(* Logix 5000 project; controller TFF vendor 1 type 14 code 107 rev 34.11; software revision 34.03 *)
// Mobius FlexReady

TASK HighPriority (periodic, rate 25 ms, priority 1, watchdog 2000 ms) : MainProgram   // High Priority Task
TASK MainTask (continuous, watchdog 500 ms) : Process, CCPSystem
TASK Task5ms (periodic, rate 5 ms, priority 10, watchdog 500 ms) : MainProgram5ms

MODULES
   Local : vendor 1 type 14 code 107 (Compact 0, rev 34.11)
      RACK_MURR_NODE1_TF3S : ETHERNET-MODULE (Ethernet 10.20.56.124, rev 1.1, Output RPI 5 ms)
      RACK_MURR_NODE5_TANK100 : ETHERNET-MODULE (Ethernet 10.20.56.162, rev 1.1, Output RPI 10 ms)
      RACK_MURR_NODE7_IND131_WI101 : ETHERNET-MODULE (Ethernet 10.20.56.141, rev 1.1, Output RPI 50 ms)
           RACK_MURR_NODE7_IND131_WI101:I.Data[1].15   // Data OK
           RACK_MURR_NODE7_IND131_WI101:I.Data[1]   // Slot 1 Scale Status
           RACK_MURR_NODE7_IND131_WI101:I.Data[0]   // Slot 1 Weight Data
           RACK_MURR_NODE7_IND131_WI101:O.Data[0]   // Slot 1 Tare/Target Value
           RACK_MURR_NODE7_IND131_WI101:O.Data[1]   // IND131 Command word Select weight display in net mode Clear all cmd excepted Tare and zero
      RACK_MURR_NODE0_SMART : ETHERNET-MODULE (Ethernet 10.20.56.131, rev 1.1, Output RPI 10 ms)
      RACK_MURR_NODE1_TF2S : ETHERNET-MODULE (Ethernet 10.20.56.123, rev 1.1, Output RPI 5 ms)
      RACK_MURR_NODE3_PUMP : ETHERNET-MODULE (Ethernet 10.20.56.151, rev 1.1, Output RPI 10 ms)
      RACK_MURR_NODE4_INSTRUM_TFF1 : ETHERNET-MODULE (Ethernet 10.20.56.172, rev 1.1, Output RPI 10 ms)
      RACK_MURR_NODE4_INSTRUM_TFF2 : ETHERNET-MODULE (Ethernet 10.20.56.173, rev 1.1, Output RPI 10 ms)
      RACK_MURR_NODE4_INSTRUM_TFF3 : ETHERNET-MODULE (Ethernet 10.20.56.174, rev 1.1, Output RPI 10 ms)
      RACK_MURR_NODE4_INSTRUM_TFF4 : ETHERNET-MODULE (Ethernet 10.20.56.175, rev 1.1, Output RPI 10 ms)
      RACK_MURR_NODE4_INSTRUM_TFF5 : ETHERNET-MODULE (Ethernet 10.20.56.176, rev 1.1, Output RPI 10 ms)
      RACK_MURR_NODE5_TANK250 : ETHERNET-MODULE (Ethernet 10.20.56.163, rev 1.1, Output RPI 10 ms)
      RACK_MURR_NODE5_TANK50 : ETHERNET-MODULE (Ethernet 10.20.56.161, rev 1.1, Output RPI 10 ms)
      RACK_MURR_NODE6_IND331_WI001 : ETHERNET-MODULE (Ethernet 10.20.56.142, rev 1.1, Output RPI 50 ms)
           RACK_MURR_NODE6_IND331_WI001:I.Data[1].15   // Data OK
           RACK_MURR_NODE6_IND331_WI001:I.Data[1]   // Slot 1 Scale Status
           RACK_MURR_NODE6_IND331_WI001:I.Data[0]   // Slot 1 Weight Data
           RACK_MURR_NODE6_IND331_WI001:O.Data[0]   // Slot 1 Tare/Target Value
           RACK_MURR_NODE6_IND331_WI001:O.Data[1]   // IND331 Command word Select weight display in net mode Clear all cmd excepted Tare and zero
END_MODULES

TYPE AlarmAnalog :   // Analog Alarm UDT
STRUCT
   Override : BOOL;   // Alarm Override
   Disable : BOOL;   // Alarm Disabled
   LOLOAlarm : BOOL;   // LOLO Alarm Condition
   LOAlarm : BOOL;   // LO Alarm Condition
   HIAlarm : BOOL;   // HI Alarm Condition
   HIHIAlarm : BOOL;   // HIHI Alarm Condition
   LOLODisable : BOOL;   // LOLO Alarm Disable
   LODisable : BOOL;   // LO Alarm Disable
   HIDisable : BOOL;   // HI Alarm Disable
   HIHIDisable : BOOL;   // HIHI Alarm Disable
   LOLOAck : BOOL;   // LOLO Alarm Acknowledged
   LOAck : BOOL;   // LO Alarm Acknowledged
   HIAck : BOOL;   // HI Alarm Acknowledged
   HIHIAck : BOOL;   // HIHI Alarm Acknowledged
   HIHIEnable : BOOL;   // HIHI Alarm Always Enabled for Critical Safety Alarms
   FeedPumpEnable : BOOL;   // LOLO and LO Alarm conditionned on Feed Pump Enable
   TransferPumpEnable : BOOL;   // LOLO and LO Alarm conditionned on Transfer Pump Enable
   LOLOAlarmONS : BOOL;   // Saves last value of alarm
   LOAlarmONS : BOOL;   // Saves last value of alarm
   HIAlarmONS : BOOL;   // Saves last value of alarm
   HIHIAlarmONS : BOOL;   // Saves last value of alarm
   FeedPumpTag : DINT;   // Feed Pump Tag for Pump Enable function
   TransferPumpTag : DINT;   // Transfer Pump Tag for Pump Enable function
   Value : DINT;   // Alarm Value : 0= No Alarm. 1=Non-Critical. 2= Non-Critical Unacknowledged. 3=Critical. 4=Critical Unacknowledged.
   ValueHMI : DINT;   // Alarm Value for HMI: 0= No Alarm. 1=Non-Critical. 2= Non-Critical Unacknowledged. 3=Critical. 4=Critical Unacknowledged.
   LOLO : REAL;   // LOLO Alarm Set Point
   LO : REAL;   // LO Alarm Set Point
   HI : REAL;   // HI Alarm Set Point
   HIHI : REAL;   // HIHI Alarm Set Point
   PV : REAL;   // Process Variable Value
   LOLOTimer : TIMER;   // LOLO Alarm Timer
   LOLOTimerSP : DINT;   // LOLO Alarm Timer setpoint (sec)
   LOTimer : TIMER;   // LO Alarm Timer
   LOTimerSP : DINT;   // LO Alarm Timer setpoint (sec)
   HITimer : TIMER;   // HI Alarm Timer
   HITimerSP : DINT;   // HI Alarm Timer setpoint (sec)
   HIHITimer : TIMER;   // HIHI Alarm Timer
   HIHITimerSP : DINT;   // HIHI Alarm Timer setpoint (sec)
   EnableCfg : BOOL;   // Set to 1 to Configure \ Use Analog Alarm
END_STRUCT
END_TYPE

TYPE AlarmControl :   // Alarm Control UDT
STRUCT
   DESC : STRING25;   // Description
   EGU : STRING5;   // Unit
   AlarmAck : BOOL;   // Alarm Acknowledge Flag
   AlarmHigh : BOOL;   // Critical Alarm Condition
   AlarmLow : BOOL;   // Non-Critical Alarm Condition
   AlarmHighUnack : BOOL;   // Critical Unacknowledged Alarm Condition
   AlarmLowUnack : BOOL;   // Non-Critical Unacknowledged Alarm Condition
   HighHMI : BOOL;   // Critical Alarm Condition (for HMI)
   LowHMI : BOOL;   // Non-Critical Alarm Condition (for HMI)
   HighUnackHMI : BOOL;   // Critical Unacknowledged Alarm Condition (for HMI)
   LowUnackHMI : BOOL;   // Non-Critical Unacknowledged Alarm Condition (for HMI)
   Horn : BOOL;   // Alarm Horn
   YellowLamp : BOOL;   // Non-Critical Alarm Indicator
   RedLamp : BOOL;   // Critical Alarm Indicator
   Current : BOOL;   // Current Alarm Status
   AckOutput : BOOL;   // Alarm Acknowledge Output
   FlashControl : BOOL;   // Flash Control
   EnableAllIn : BOOL;   // Enable All Alarms Input
   EnableAllOut : BOOL;   // Enable All Alarms Output
   DisableAllIn : BOOL;   // Disable All Alarms Input
   DisableAllOut : BOOL;   // Disable All Alarms Output
   NewAlarm : BOOL;   // True for 1 scan when new alarm is detected
   SilenceHorn : BOOL;   // Set true to Silence horn
   FlashTimer : TIMER;   // Flash Timer
   AckTimer : TIMER;   // Acknowledge Timer
   EnableAllTimer : TIMER;   // Enable All Alarms Timer
   DisableAllTimer : TIMER;   // Disable All Alarms Timer
   HornAddress : INT;   // Output address for Alarm horn
   EnableAllAnaSigIn : BOOL;   // Enable All analog signal failure Alarms Input
   EnableAllAnaSigOut : BOOL;   // Enable All analog signal failure Alarms Output
   DisableAllAnaSigIn : BOOL;   // Disable All analog signal failure Alarms Input
   DisableAllAnaSigOut : BOOL;   // Disable All analog signal failure Alarms Output
   EnableAllAnaSigTimer : TIMER;   // Enable All analog signal failure Alarms Timer
   DisableAllAnaSigTimer : TIMER;   // Disable All analog signal failure Alarms Timer
   AlarmHighMem : BOOL;   // Critical Alarm Condition Mem
   ESAckAddress : INT;   // Output address for re-established system
   ESAckTimer : TIMER;   // Emergency Stop Acknowledge Timer
   ESAck : BOOL;   // Emergency Stop Acknowledge
   InitAlarmConfig : BOOL;   // Initialize alarms config if the command is set from the HMI
END_STRUCT
END_TYPE

TYPE AlarmDeviation :   // Deviation Alarm UDT
STRUCT
   Override : BOOL;   // Alarm Override
   Disable : BOOL;   // Alarm Disabled
   HIAlarm : BOOL;   // HI Deviation Alarm Condition
   HIHIAlarm : BOOL;   // HIHI Deviation Alarm Condition
   HIDisable : BOOL;   // HI Alarm Disable
   HIHIDisable : BOOL;   // HIHI Alarm Disable
   HIAck : BOOL;   // HI Alarm Acknowledged
   HIHIAck : BOOL;   // HIHI Alarm Acknowledged
   LOLOAlarmONS : BOOL;   // One shot when alarm occures
   HIAlarmONS : BOOL;   // One shot when alarm occures
   LOAlarmONS : BOOL;   // One shot when alarm occures
   HIHIAlarmONS : BOOL;   // One shot when alarm occures
   Value : DINT;   // Alarm Value
   ValueHMI : DINT;   // Alarm Value for HMI
   HI : REAL;   // HI Alarm Set Point
   HIHI : REAL;   // HIHI Alarm Set Point
   LOLOLim : REAL;   // LOLO Alarm Set Point (calculated)
   LOLim : REAL;   // LO Alarm Set Point (calculated)
   HILim : REAL;   // HI Alarm Set Point (calculated)
   HIHILim : REAL;   // HIHI Alarm Set Point (calculated)
   HITimer : TIMER;   // HI Alarm Timer
   HITimerSP : DINT;   // HI Alarm Timer setpoint (sec)
   HIHITimer : TIMER;   // HIHI Alarm Timer
   HIHITImerSP : DINT;   // HIHI Alarm Timer setpoint (sec)
   EnableCfg : BOOL;   // Set to enable alarm
END_STRUCT
END_TYPE

TYPE AnalogInput :   // Analog Input UDT
STRUCT
   TagName : STRING6;   // PID Tag Name
   TagDisplayName : STRING6;   // PID Tag Name
   OutofRange : BOOL;   // Out of Range
   FilterType : BOOL;   // Filter Type 0=LP, 1=Avg
   AveragingTotal : DINT;   // Averaging Filter Total
   Address : DINT;   // Input Address (RawAnalogInputArray)
   RawMin : DINT;   // Raw Minimum Range
   RawMax : DINT;   // Raw Maximum Range
   RawValue : DINT;   // Raw Value (Measuring value given by the I/O card)
   RawLowLimit : DINT;   // Raw Out of Range LO Limit
   RawHighLimit : DINT;   // Raw Out of Range HI Limit
   FilterUser : DINT;   // User Filter Value
   FilteredRaw : DINT;   // Raw Filtered Value
   FilterActual : REAL;   // Actual Filter Value
   ScaledMin : REAL;   // Scaled Minimum Range
   ScaledMax : REAL;   // Scaled Maximum Range
   CurrentValue : REAL;   // Current Value
   RangeMin : REAL;   // Scaled Minimum Range (Config Analog Points)
   RangeMax : REAL;   // Scaled Maximum Range (Config Analog Points)
   RangeMinSave : REAL;   // Scaled Minimum Range (previous)
   RangeMaxSave : REAL;   // Scaled Maximum Range (previous)
   RealCfg : BOOL;   // Set to 1 if real analog input is used. Set to 0 for soft input (derived data)
   EnableCfg : BOOL;   // Set to 1 to activate this Tag
   OverrideCfg : BOOL;   // Set to 1 to allow user to Overide alarm
   Desc : STRING25;   // Description
   EGU : STRING5;   // Unit
END_STRUCT
END_TYPE

TYPE AnalogOutput :   // Analog Output UDT
STRUCT
   Tag : STRING10;   // Tag name
   RawValue : DINT;   // Raw Value Send to I/O Card
   RawMin : DINT;   // Raw Min
   RawMax : DINT;   // Raw Max
   ScaledValue : REAL;   // Scaled Value
   ScaledMin : REAL;   // Scaled Minimum Range
   ScaledMax : REAL;   // Scaled Maximum Range
   EnableCfg : BOOL;   // Set to 1 to enable Analog Output
END_STRUCT
END_TYPE

TYPE AverageCalculation :
STRUCT
   SUM : REAL;   // Sum of average
   COUNTER : DINT;   // Counter of average
   TIMER : TIMER;   // Timer of average
   TIMER_OSR : BOOL;   // Timer one shot
END_STRUCT
END_TYPE

TYPE CCPSystem :   // CCP System UDT
STRUCT
   Run : BOOL;   // Run Flag
   RunAuto : BOOL;   // Auto Run Flag
   Procedure : BOOL;   // Procedure Flag
   Complete : BOOL;   // Procedure Complete
   Download : BOOL;   // Manual Download
   Heartbeat : BOOL;   // CCPRuntime Heartbeat
   OperationDownloadFlag : BOOL;   // Legacy Tag. Not used by PLC
   OperationStartFlag : BOOL;   // Operation Start Flag
   Manual : BOOL;   // Recipe Pool Flag
   State : DINT;   // Machine State
   Language : DINT;   // Language Number
   ErrorPhase : DINT;   // Error in Phase #
   ErrorStep : DINT;   // Error in Step #
   Error : DINT;   // Error Description
   OperationNoInBatch : DINT;   // Legacy Tag. Not used by PLC
   EndPointer : DINT;   // End Operation Step Buffer Pointer
   Machine : STRING;   // Machine Name
   ProductID : STRING;   // Batch Product ID from Operation Header
   Description : STRING;   // Batch Description from Operation Header
   Created : STRING;   // Date and Time when the last operation has been downloaded in PLC
   Originator : STRING;   // Last saved by field from Operation Header
   Comment : STRING;   // Comment
   OperationName : STRING90;   // Name and path of last operation downloaded in PLC
   ConfigFile : STRING;   // Current configuration file used
   LastMod : STRING;   // Last Mod
   GradientBasis : STRING;   // Gradient Basis
   GradientVariable : STRING;   // Gradient Variable
   GradientSegments : STRING;   // Gradient Segments
   StateWatchDog : TIMER;   // If Downloading for longer than this time the state will reset to 0
   EventList : EventList;   // Event List Array
   BufferSteps : STRING25[251];   // Buffer Steps Array
   BufferEvents : STRING50[251];   // Buffer Events Array
   HETP_ON_OFF : BOOL;   // HETP (1 = Start , 0 = Stop)
   DefaultOnComplete : BOOL;   // At the end of recipe apply default flowpath (0 = Apply , 1 = Don't Apply)
END_STRUCT
END_TYPE

TYPE CCPSystem_Storage :
STRUCT
   Run : BOOL;   // Run Flag
   RunAuto : BOOL;   // Auto Run Flag
   Procedure : BOOL;   // Procedure Flag
   Complete : BOOL;   // Procedure Complete
   Download : BOOL;   // Manual Download
   Heartbeat : BOOL;   // CCPRuntime Heartbeat
   OperationDownloadFlag : BOOL;   // Legacy Tag. Not used by PLC
   OperationStartFlag : BOOL;   // Operation Start Flag
   TestAction : BOOL;   // Action Test Flag
   Manual : BOOL;   // Recipe Pool Flag
   State : DINT;   // Machine State
   Language : DINT;   // Language Number
   ErrorPhase : DINT;   // Error in Phase #
   ErrorStep : DINT;   // Error in Step #
   Error : DINT;   // Error Description
   OperationNoInBatch : DINT;   // Legacy Tag. Not used by PLC
   EndPointer : DINT;   // End Operation Step Buffer Pointer
   Machine : STRING;
   ProductID : STRING;
   Description : STRING;
   Created : STRING;
   Originator : STRING;
   Comment : STRING;
   OperationName : STRING90;
   ConfigFile : STRING;
   LastMod : STRING;
   GradientBasis : STRING;
   GradientVariable : STRING;
   GradientSegments : STRING;
   StateWatchDog : TIMER;   // If Downloading for longer than this time the state will reset to 0
END_STRUCT
END_TYPE

TYPE ChartMark :   // Chart Mark UDT
STRUCT
   In : BOOL;   // Chart Mark In
   Out : BOOL;   // Chart Mark Out
END_STRUCT
END_TYPE

TYPE Concentration :   // Concentration UDT
STRUCT
   VCF : REAL;   // Volume Concentration Factor
   CB : REAL;   // Protein Concentration
   Conc_Init : REAL;   // Initial Protein Concentration SP
   Conc_Final : REAL;   // Final Protein Concentration SP
   Conc_Final_Volume : REAL;   // Final Concentration Volume SP
   Final_Conc_Volume_Reached : BOOL;   // Final Concentration Volume Reached
   Final_Conc_Volume_DownTimer : TIMER;   // Final Concentration Volume Deactivation timer
   Final_Conc_Volume_UpTimer : TIMER;   // Final Concentration Volume Activation timer
   Final_Conc_Protein_Reached : BOOL;   // Final Protein Concentration Reached
   Final_Conc_Protein_DownTimer : TIMER;   // Final Protein Concentration Deactivation timer
   Final_Conc_Protein_UpTimer : TIMER;   // Final Protein Concentration Activation timer
   LogConcIn : BOOL;   // Log Concentration Input
   LogConcOut : BOOL;   // Log Concentration Output
   LogConcTimer : TIMER;   // Log Concentation Timer
END_STRUCT
END_TYPE

TYPE Configuration :   // Configuration UDT
STRUCT
   Reset : BOOL;   // Activate Reset Loop Configuration
   IndexA0 : DINT;   // Index AnalogOutput
   IndexAP : DINT;   // Index AnalogPoint
   IndexDP : DINT;   // Index DigitalPoint
   IndexDr : DINT;   // Index Drive
   IndeXValve : DINT;   // Index Valve
   IndexReset : DINT;   // Index Reset
   IndexCL : DINT;   // Index Control Loop
   IndexFlowpath : DINT;   // Index Flowpath
END_STRUCT
END_TYPE

TYPE ControlLoop :   // Control Loop UDT
STRUCT
   Tag : STRING5;   // Tag Name
   Desc : STRING25;   // Description
   LoopCfg : BOOL;   // Set to 1 to use this loop
   ManualEGU : STRING5;   // Unit of Manual Control Mode
   AutoEGU : STRING5;   // Unit of Auto Control Mode
   Auto1EGU : STRING5;   // Unit of Auto Control Mode 1
   Auto2EGU : STRING5;   // Unit of Auto Control Mode 2
   Auto3EGU : STRING5;   // Unit of Auto Control Mode 3
   Interlock : BOOL;   // Loop Interlock
   Enable : BOOL;   // Loop Enabled
   Manual : BOOL;   // Control Mode 0=Auto, 1=Manual
   Stable : BOOL;   // Loop Stable
   DBOK : BOOL;   // Control Within Deadband
   Status : INT;   // Status
   Auto1 : BOOL;   // Auto Control Mode 1
   Auto2 : BOOL;   // Auto Control Mode 2
   Auto3 : BOOL;   // Auto Control Mode 3
   Auto4 : BOOL;   // Auto Control Mode 4
   StepUp : BOOL;   // Increment CV
   StepDown : BOOL;   // Decrement CV
   RampEnable : BOOL;   // Ramp Enable
   RampUp : BOOL;   // Ramping UP
   RampDown : BOOL;   // Ramping Down
   RampStatus : BOOL;   // Ramping Status
   RampAutoOSR : BOOL;   // Auto Ramp One-Shot
   RampManualOSR : BOOL;   // Manual Ramp One-Shot
   PIDEnable : BOOL;   // PID Enabled
   ManualOSR : BOOL;   // Manual Mode One-Shot
   Auto1OSR : BOOL;   // Control Mode 1 One-Shot
   Auto2OSR : BOOL;   // Control Mode 2 One-Shot
   Auto3OSR : BOOL;   // Control Mode 3 One-Shot
   Auto4OSR : BOOL;   // Control Mode 4 One-Shot
   StepIncrement : DINT;   // Step Increment/Decrement Value
   CycleTime : DINT;   // Cycle Time (for modulating output)
   PV : REAL;   // Process Variable
   PVAuto1 : REAL;   // Process Variable for Control Mode Auto 1
   PVAuto2 : REAL;   // Process Variable for Control Mode Auto 2
   PVAuto3 : REAL;   // Process Variable for Control Mode Auto 3
   PVAuto4 : REAL;   // Process Variable for Control Mode Auto 4
   CV : REAL;   // Control Value
   SPAuto : REAL;   // Auto Set Point
   SPAutoSave : REAL;   // Auto Set Point (previous)
   SPAuto1 : REAL;   // Auto Set Point Mode 1
   SPAuto2 : REAL;   // Auto Set Point Mode 2
   SPAuto3 : REAL;   // Auto Set Point Mode 3
   SPAuto4 : REAL;   // Auto Set Point Mode 4
   SPManual : REAL;   // Manual Set Point
   SPManualSave : REAL;   // Manual Set Point (previous)
   RangeMin : REAL;   // Min EGU Range
   RangeMax : REAL;   // Max EGU Range
   SPRangeMin : REAL;   // Set Point Min EGU Range
   SPRangeMax : REAL;   // Set Point Max EGU Range
   RampRate : REAL;   // Ramp Rate
   RampRateSave : REAL;   // Ramp Rate (previous)
   RampStart : REAL;   // Ramp Start Value
   Deadband : REAL;   // Deadband
   DBLO : REAL;   // Low Deadband Value
   DBHI : REAL;   // High Deadband Value
   RampTimer : TIMER;   // Ramp Timer
   StableTimer : TIMER;   // Loop Stable Timer
   StableTime : DINT;   // Loop Stable Time setpoint (sec)
   PIDTimer : TIMER;   // PID Timer
   CycleTimer : TIMER;   // Cycle Timer (for modulating output)
   PID : PID;   // PID Instruction Data
   KP : REAL[3];   // Loop Gain from HMI
   KI : REAL[3];   // Loop Reset from HMI
   KD : REAL[3];   // Loop Rate from HMI
   DB : REAL[3];   // Loop Deadband from HMI
   On : BOOL;   // Turns all controll On
   DisOSR : BOOL;   // One Shot DisOSR
   OutputOn_OSR : BOOL;   // One Shot OutputOn_OSR
   OutputOff_OSR : BOOL;   // One Shot OutputOff_OSR
   DigitalOutput : BOOL;   // Output from loop in for descrete control
   RampCfg : BOOL;   // Set to 1 to Enable Ramp Option
   Auto1Cfg : BOOL;   // Set to 1 to use Auto 1 option
   Auto2Cfg : BOOL;   // Set to 1 to use Auto 2 option
   Auto3Cfg : BOOL;   // Set to 1 to use Auto 3 option
   Auto4Cfg : BOOL;   // Set to 1 to use Auto 4 option
   Auto1PVCfg : DINT;   // Set to Analog Point Number
   Auto2PVCfg : DINT;   // Set to Analog Point Number
   Auto3PVCfg : DINT;   // Set to Analog Point Number
   Auto4PVCfg : DINT;   // Set to Analog Point Number
   Auto1RangeMax : REAL;   // Set Point EGU Range Max
   Auto2RangeMax : REAL;   // Set Point EGU Range Max
   Auto3RangeMax : REAL;   // Set Point EGU Range Max
   Auto4RangeMax : REAL;   // Set Point EGU Range Max
   AutoSwitchEnable : BOOL;   // Set to 1 to allow loop to switch from auto1 to auto 2
   OutputAddress : INT;   // Set to analog output to use for this loop
   LoopStatus : INT;   // Loop Mode Status for HMI
END_STRUCT
END_TYPE

TYPE CriteriaFlag :   // Criteria Flag UDT
STRUCT
   Flag1 : BOOL;   // Criteria Flag 1 (1=ON , 0=OFF)
   Flag2 : BOOL;   // Criteria Flag 2 (1=ON , 0=OFF)
   Flag3 : BOOL;   // Criteria Flag 3 (1=ON , 0=OFF)
   Flag4 : BOOL;   // Criteria Flag 4 (1=ON , 0=OFF)
   Flag5 : BOOL;   // Criteria Flag 5 (1=ON , 0=OFF)
END_STRUCT
END_TYPE

TYPE CVTune :   // Control Valve Tuning Data Type
STRUCT
   ClosedRaw : REAL;   // Captured Raw Value When Valve is Closed
   OpenRaw : REAL;   // Captured Raw Value When Valve is Open
   MinOutput : REAL;   // Minimum output for tuning adjustment for valve
   MaxOutput : REAL;   // Maximum output for tuning adjustment for valve
   MinTimer : TIMER;   // Timer to capture closed raw value
   MaxTimer : TIMER;   // Timer to capture open raw value
   OSR : INT;   // One shot bits
   Activate : BOOL;   // Activate tuning function
   Enable : BOOL;   // Tuning routine is enabled
END_STRUCT
END_TYPE

TYPE DCS :
STRUCT
   ActionsParameters : DCSParameters;   // Recipe Parameters
   Criteria : DCSCriteria;   // Recipe Criteria
   RunCmd : BOOL;   // Start Recipe Command
   ShowHeader : BOOL;   // Show Pre and Post Run Header
   RunID : STRING50;   // Recipe Header Run ID (Must be unique)
   UserName : STRING80;   // Recipe Header User Name
   ProductID : STRING80;   // Recipe Header Product ID
   BatchID : STRING80;   // Recipe Header Batch ID
   StepID : STRING80;   // Recipe Header Step ID
   FileName : STRING240;   // File Name for Start recipe (if not using RecipePoolID)
   PreRunComment : STRING240;   // Recipe Header Pre Run Comment
   PostRunComment : STRING240;   // Recipe Header Post Run Comment
   RecipePoolID : DINT;   // Recipe Pool ID for Start recipe (If 0 the file name will be used)
   Status : DINT;   // System status for DCS
   ColumnInfo : STRING240;   // Recipe Header Column Info
   PackedBedInfo : STRING240;   // Recipe Header Packed Bed Info
   SampleInfo : STRING240;   // Recipe Header Sample Info
   BufferInfo : STRING240;   // Recipe Header Buffer Info
END_STRUCT
END_TYPE

TYPE DCSCriteria :
STRUCT
   Criteria_1 : BOOL;
   Criteria_2 : BOOL;
END_STRUCT
END_TYPE

TYPE DCSParameters :
STRUCT
   Feed_Pump_Speed_Setpoint : REAL[3];
   Feed_Pump_Flow_Setpoint : REAL[3];
   Feed_Pump_DP_Setpoint : REAL[3];
   Level_Pump_Speed_Setpoint : REAL[3];
   Level_Pump_Level_Setpoint : REAL[3];
   PCV001_Retentate_Position_Setpoint : REAL[3];
   PCV001_Retentate_Pressure_Setpoint : REAL[3];
   PCV001_Retentate_TMP_Setpoint : REAL[3];
   PCV101_Filtrate_Position_Setpoint : REAL[3];
   PCV101_Filtrate_Flow_Setpoint : REAL[3];
   PCV101_Filtrate_TMP_Setpoint : REAL[3];
   Mixer_Speed_Setpoint : REAL[3];
   Mixer_Auto_Min_Setpoint : REAL[3];
   Mixer_Auto_Max_Setpoint : REAL[3];
   Init_Protein_Conc : REAL[1];
   Final_Protein_Conc : REAL[1];
   Final_Protein_Volume : REAL[1];
   Holdup_Volume : REAL[1];
   Init_Diaf_Volume : REAL[1];
   Final_Diaf_Volume : REAL[1];
   Membrane_Area : REAL[1];
   Membrane_Density : REAL[1];
END_STRUCT
END_TYPE

TYPE DerivedData :   // DerivedData UDT
STRUCT
   HOLDUP : REAL;   // Holdup Volume
   PI001_PSI : REAL;   // PI001 Pressure in PSI
   PI401_PSI : REAL;   // PI401 Pressure in PSI
END_STRUCT
END_TYPE

TYPE Diafiltration :   // Diafiltration UDT
STRUCT
   Diaf_Volume : REAL;   // Diafiltration Volume
   Diaf_Init : REAL;   // Initial Diafiltration Volume SP
   Diaf_Final_Volume : REAL;   // Final Diafiltration Volume SP
   Snap : BOOL;   // Level Snapshot
   Final_Diaf_Volum_Reached : BOOL;   // Final Diafiltration Volume Reached
   Final_Diaf_Volum_DownTimer : TIMER;   // Final Diafiltration Volume Deactivation timer
   Final_Diaf_Volum_UpTimer : TIMER;   // Final Diafiltration Volume Activation timer
   Diaf_Snap_Value : REAL;   // Volume value snapped
   LogDiafIn : BOOL;   // Log Diafiltration Input
   LogDiafOut : BOOL;   // Log Diafiltration Output
   LogDiafTimer : TIMER;   // Log Diafiltration Timer
END_STRUCT
END_TYPE

TYPE DigitalPoint :   // Digital Point UDT
STRUCT
   Tag : STRING10;   // PID Tag to be Used for Display
   Desc : STRING25;   // Description to be Used for Display
   CurrentValue : BOOL;   // Current value of Tag
   AlarmCurrentValue : BOOL;   // Displays state of processed alarm input.
   AlarmAck : BOOL;   // Alarm Acknowledged
   Alarm : BOOL;   // Alarm
   Override : BOOL;   // Alarm Override
   Mimic : INT;   // Set color on HMI digital point mimic
   SoftInput : BOOL;   // Used as current value when RealInputCfg is set to 0
   Condition1 : BOOL;   // Enable Condition 1 Must be True to Enable alarm condition
   Condition2 : BOOL;   // Enable Condition 2 Must be True to Enable alarm condition
   Cond1Text : STRING;   // Condtion 1 Text
   Cond2Text : STRING;   // Condition 2 text
   DelayTimer : TIMER;   // Alarm Timer
   DelayTimerSP : DINT;   // Alarm Timer setpoint (sec)
   Priority : BOOL;   // Alarm Priority 0=Low, 1=High
   EnableCfg : BOOL;   // Set to True to configure point on system
   ActiveStateCFg : BOOL;   // Set to 0 to invert incomming state
   RealInputCfg : BOOL;   // Set to 1 to Use Hardwired Input. Set to 0 to disable Hardwired and use software condition
   InputAddressCfg : DINT;   // Set to address of hardwared input to be used on alarm
   AlarmCfg : BOOL;   // Set to 1 to Use alarm on this point
   AlarmStateCfg : BOOL;   // Set to 1 to alarm on a 0 to 1 transition. Set to zero to alarm on a 1 to 0 transition
   OverrideCfg : BOOL;   // set to 1 to allow user to Override alarm
   PriorityCfg : BOOL;   // Set to 1 to allow user to set Priority and Enable
   Cond1Cfg : BOOL;   // Set to 1 to Enable Condition
   Cond2Cfg : BOOL;   // Set to 1 to Enable Condition
   FlashingInputCfg : BOOL;   // Set to 1 for Heartbeat Style Inputs
   AlarmONS : BOOL;   // One shot when alarm occurs
END_STRUCT
END_TYPE

TYPE Drive :   // Pump Control UDT
STRUCT
   TagName : STRING10;   // Drive tag name
   Desc : STRING25;   // Drive Description
   Mode : BOOL;   // Control Mode
   ManualCommand : BOOL;   // Manual Command
   AutoCommand : BOOL;   // Auto Command
   RunCommand : BOOL;   // Run Command
   RunStatus : BOOL;   // Running Status
   RunInterlock : BOOL;   // Run Interlock
   RunInput : BOOL;   // Run Digital Input 0=No, 1=Yes
   OutputAddress : DINT;   // Run Command Output Address
   InputAddress : DINT;   // Running Input Address
   InterlockTimer : TIMER;   // Interlock Delay Timer
   RunOns : BOOL;   // Run one shot
   StopOns : BOOL;   // Stop One shot
   RunRequest : BOOL;   // Run request for auto or man mode
   Interlocked : BOOL;   // Drive is commanded to run but currently stopped by interlock
   EnableCfg : BOOL;   // Set to enable Drive
   ReverseCfg : BOOL;   // Set to enable reverse control
   Direction : BOOL;   // 0 = forward. 1 = reverse
   DirectionAddress : DINT;   // Direction Output Address
   DriveStatus : INT;   // Drive Status
   DriveLoopStatus : INT;   // Drive Loop Status
   DriveAlarmStatus : INT;   // Drive Alarm Status
   ValidFlowpath : BOOL;   // Valid flowpath flag
END_STRUCT
END_TYPE

TYPE EventList :
STRUCT
   Event : DINT[1000];   // Event List Array
   Value : REAL[1000];   // Value Array
   PreRunValue : REAL[1000];   // Pre Run Value
END_STRUCT
END_TYPE

TYPE FactorySettings :   // Factory Settings
STRUCT
   ProductName : STRING90;   // Product Name
   SerialNumber : STRING90;   // Serial Number
   ComputerName : STRING90;   // Computer Name
   ComputerDesc : STRING90;   // Computer Description
   DateFormat : STRING90;   // Date Format
   FlagUK : BOOL;   // Use UK Flag instead of US
   PCV001ClosedSP : REAL;   // PCV001 Closed Set Point
   PCV101ClosedSP : REAL;   // PCV101 Closed Set Point
END_STRUCT
END_TYPE

TYPE FaultRecordType :   // Fault Record Type UDT
STRUCT
   TimeLow : DINT;   // Lower 32 bits of the fault timestamp value
   TimeHigh : DINT;   // Upperer 32 bits of the fault timestamp value
   RecType : INT;   // Fault Type
   Code : INT;   // Unique code for the fault
   Info : DINT[8];   // Fault specific information
END_STRUCT
END_TYPE

TYPE FlowPath :   // Flow Path UDT
STRUCT
   Command : BOOL;   // Flow Path Command
   Status : BOOL;   // Flow Path Status
   FlushTruth : BOOL;   // Flush Mode Enable Truth
   DrainTruth : BOOL;   // Drain Mode Enable Truth
   FlushMask : BOOL;   // Flush Mode Enable Mask
   DrainMask : BOOL;   // Drain Mode Enable Mask
   Truth1 : DINT;   // Truth Table 1 (Valves 1-32)
   Truth2 : DINT;   // Truth Table 2 (Valves 33-64)
   Truth3 : DINT;   // Truth Table 3 (Valves 65-96)
   Truth4 : DINT;   // Truth Table 4 (Valves 97-128)
   Mask1 : DINT;   // Mask 1 (Valves 1-32)
   Mask2 : DINT;   // Mask 2 (Valves 33-64)
   Mask3 : DINT;   // Mask 3 (Valves 65-96)
   Mask4 : DINT;   // Mask 4 (Valves 97-128)
   Desc : STRING;   // Flow Path Description
END_STRUCT
END_TYPE

TYPE FlowPathControl :   // Flow Path Control UDT
STRUCT
   Flag : BOOL;   // Flow Path Command Flag
   Valve1 : DINT;   // Valve Control 1 (Valves 1-32)
   Valve2 : DINT;   // Valve Control 2 (Valves 33-64)
   Valve3 : DINT;   // Valve Control 3 (Valves 65-96)
   Valve4 : DINT;   // Valve Control 4 (Valves 97-128)
   MaxFlowPath : DINT;   // Maximum Number of Flow Paths
   Status : DINT;   // Flow Path Status
   StatusHMI : DINT;   // Flow Path Status for HMI
   Save : BOOL;   // Set to 1 to save Flowpath
   SaveStored : BOOL;   // Stored Save cmd
   Restore : BOOL;   // Set to 1 to restore flowpath
   SaveOns : BOOL;   // one shot after save
   HoldOns : BOOL;   // one shot after Hold
   FlowpathEnable : BOOL[64];   // Enable Flowpath
   FlushMode_Enabled : BOOL;   // Flush Mode Enabled
   DrainMode_Enabled : BOOL;   // Drain Mode Enabled
END_STRUCT
END_TYPE

TYPE FlowPathSetup :   // Flowpath Setup UDT
STRUCT
   Apply : BOOL;   // Apply Flow Path
   Number : DINT;   // Flow Path Number
   Prev : DINT;   // Previous Flow Path Number
   Mask_View : BOOL;   // View the Mask of selected Flowpath
   Mask_Save : BOOL;   // Save the Mask of selected Flowpath
   Truth_View : BOOL;   // View the Truth of selected Flowpath
   Truth_Save : BOOL;   // Save the Truth of selected Flowpath
   OpenAllValve : BOOL;   // Set the Flowpath 61 to Open All Valves
   CloseAllValve : BOOL;   // Set the Flowpath 62 to Close All Valves
END_STRUCT
END_TYPE

TYPE IO_Station :   // Station State UDT
STRUCT
   Node_Comm_Status_value : INT;   // Node Communication Status Value (get from status of hardware card)
   Node_Comm_Status : BOOL;   // Node Communication Status (0=Defect , 1=OK)
   Node_Internal_Defect_Status_value : INT;   // Node Internal Defect Status Value (at least one defect on the node : branch, slot, channel)
   Node_Internal_Defect_Status : BOOL;   // Node Internal Defect Status (0=Defect , 1=OK)
   Inhibition : DINT;   // Inhibit \ Uninhibit Station Module
END_STRUCT
END_TYPE

TYPE LinearGradient :   // Linear Gradient UDT
STRUCT
   Enable : BOOL;   // Linear Gradient Enable
   Hold : BOOL;   // Gradient Hold
   Segments : DINT;   // Number of Segments
   Variable : DINT;   // Gradient Variable (1=Time, 2=CVs, 3=Volume)
   Basis : DINT;   // Basis (1=Percent, 2=Conductivity)
   Segment : DINT;   // Current Segment
   State : DINT;   // Sets state of control : 0 = Disabled 1 = Running 2 = Paused
   Input : REAL;   // Input Value
   Result : REAL;   // Result
   X2 : REAL;   // Current Segment Duration
   Y1 : REAL;   // Current Start Value
   Y2 : REAL;   // Current End Value
   X : REAL[21];   // Gradient X Values (Durations)
   Y : REAL[21];   // Gradient Y Values (Set Points)
END_STRUCT
END_TYPE

TYPE LoggedValue :   // Logged Value UDT
STRUCT
   Value : REAL[8];   // Value to be logged in Audit Trail (used in Event section of configuration file)
END_STRUCT
END_TYPE

TYPE Membrane_Data :   // Membrane Data UDT
STRUCT
   Flux : REAL;   // Membrane Flux
   Area : REAL;   // Membrane Area SP
   Density : REAL;   // Density
   NWP_TCF : REAL;   // NWP Temperature correction factor
   NWP_TCF_Temp : INT;   // Temp. Temperature used in NWP calculation (INT)
   NWP_TCF_Lookup_25 : REAL[53];   // Lookup table for TCF
   AlarmStatus : INT;   // Alarm Status ( 0 = No Alarm , 1 = Non Critical Alarm , 2 = Critical Alarm )
END_STRUCT
END_TYPE

TYPE Memory_Data :   // This UDT is for putting the memory information returned by the Controller
STRUCT
   Reading_Request : BOOL;   // Request of Memory data reading
   Free_Mem_IO : DINT;   // Controler data: Free I/O Memory
   Free_Mem_DT : DINT;   // Controler data: Free Data & Logic Memory
   Free_Mem_Gen : DINT;   // Controler 1756-L55M16 only: Free Expansion Memory
   Free_Memory : DINT;   // Controler data: Total Free Memory (addition)
   Total_Mem_IO : DINT;   // Controler data: Total I/O Memory
   Total_Mem_DT : DINT;   // Controler data: Total Data & Logic Memory
   Total_Mem_Gen : DINT;   // Controler 1756-L55M16 only: Total Expansion Memory
   Total_Memory : DINT;   // Controler data: Total Memory (addition)
   Biggest_Gen_Mem_Size_Ava : DINT;   // Controler 1756-L55M16 only: Additionnal Expansion Memory
   Biggest_IO_Mem_Size_Ava : DINT;   // Controler 1756-L55M16 only: Largest contiguous block of Additionnal free Expansion Memory
   Biggest_DT_Mem_Size_Ava : DINT;   // Controler dsata: Largest contiguous block of Additionnal free Expansion Memory
   Total_Mem_DT_Real : REAL;   // Controler data: Total Data & Logic Memory
   Free_Mem_DT_Real : REAL;   // Controler data: Free Data & Logic Memory
   Used_Mem_DT_Real : REAL;   // Controler data: Used Data & Logic Memory
   Percentage_Used_DT : REAL;   // Controler data: Percentage of used Data & Logic Memory
END_STRUCT
END_TYPE

TYPE Mixer :
STRUCT
   Enable : BOOL;   // Enable Mixer Control Loop
   Mode : BOOL;   // Control Mode 0=Weight, 1=Speed
   ModeONS : BOOL;   // Manual Mode One-Shot
   SPManual : REAL;   // Manual Speed Set Point
   SPAutoMin : REAL;   // Auto Max Speed Set Point
   SPAutoMax : REAL;   // Auto Min Speed Set Point
   LevelMin : REAL;   // Minimum Level
   LevelMax : REAL;   // Maximum Level
   CV : REAL;   // Control Value
   Alarm_Reset_Cmd : BOOL;   // Alarm Reset Command
   Alarm_Reset_Cmd_Timer : TIMER;   // Alarm Reset Command Timer
END_STRUCT
END_TYPE

TYPE OperatingTime :   // Operating Time Exceeded Control
STRUCT
   DayMax : REAL;   // Setpoint for Alarm Operating Time Exceeded
   HMICtrl : BOOL;   // Control Tag Reset on launch Workspace
   TimerCtrl : TIMER;   // Timer for set tag HMICtrl
   CountPre : DINT;   // Setpoint for Alarm in sec
   Counter : DINT;   // Second Counter for Alarm
END_STRUCT
END_TYPE

TYPE Operation :   // Operation UDT
STRUCT
   Step : DINT;   // Step Number
   Criteria1 : DINT;   // Criteria 1 Code
   Criteria1Operator : DINT;   // Criteria 1 Operator
   Boolean : DINT;   // Boolean
   Criteria2 : DINT;   // Criteria 2 Code
   Criteria2Operator : DINT;   // Criteria 2 Operator
   Action : DINT;   // Action Code
   Label : DINT;   // Label
   Criteria1Value : REAL;   // Criteria 1 Value
   Criteria2Value : REAL;   // Criteria 2 Value
   ActionValue : REAL;   // Action Value
END_STRUCT
END_TYPE

TYPE Options :   // Options UDT
STRUCT
   No_Filtrate_Measurement : BOOL;   // No Filtrate Measurement
   WI101 : BOOL;   // WI101 Filtrate Weight
   WI102 : BOOL;   // WI102 Customer Filtrate Weight
   FI101 : BOOL;   // FI101 Filtrate Flow Meter
   WI101_FI101 : BOOL;   // WI101 Filtrate Weight + FI101 Filtrate Flow Meter
   WI102_FI101 : BOOL;   // WI102 Customer Filtrate Weight + FI101 Filtrate Flow Meter
   No_Device_Connected : BOOL;   // No Device Connected
   AI102_AI103 : BOOL;   // Instrum TFF1 : AI102 + AI103
   AI101 : BOOL;   // Instrum TFF2 : AI101
   AI101_AI102_AI103 : BOOL;   // Instrum TFF3 : AI101 + AI102 + AI103
   AI101_AI104 : BOOL;   // Instrum TFF4 : AI101 + AI104
   AI101_AI102_AI103_AI104 : BOOL;   // Instrum TFF5 : AI101 + AI102 + AI103 + AI104
   No_Tank : BOOL;   // No Tank connected
   Tank50 : BOOL;   // Tank 50L
   Tank100 : BOOL;   // Tank 100L
   Tank250 : BOOL;   // Tank 250L
   CCP_Report : BOOL;   // CCP Report
   TF2S : BOOL;   // TF2S installed
   TF3S : BOOL;   // TF3S installed
   ClosedFP : BOOL;   // Fully Closed Flowpath custom option
   FI003 : BOOL;   // Retentate Flowmeter custom option
END_STRUCT
END_TYPE

TYPE PCV :
STRUCT
   SP : REAL;
   PV : REAL;
   ERREUR : REAL;
   CV : REAL;
   KP : REAL;
   KI : REAL;
   TP : REAL;
   TI : REAL;
   ACCU_TI : REAL;
   OpenRawValue : REAL;
   ClosedRawValue : REAL;
   RESET : BOOL;
END_STRUCT
END_TYPE

TYPE PCV_Calib :   // PCV Position Calibration
STRUCT
   Activate : BOOL;   // Calibration Command from HMI
   Enable : BOOL;   // PCV Calibration function enabled
   OSR : INT;   // One Shot bits
   Open_SP_Target : REAL;   // Open setpoint of PCV to achieve
   Close_SP_Target : REAL;   // Close setpoint of PCV to achieve
   Open_Timer : TIMER;   // Timer before save the raw value
   Close_Timer : TIMER;   // Timer before save the raw value
END_STRUCT
END_TYPE

TYPE PCV_Control :   // PCV Control UDT
STRUCT
   FullOpen : BOOL;   // fully open the valve without ramp
   FullOpenSP : REAL;   // target value of the valve opening
   FullOpenResetTimer : TIMER;   // Timer to reset full open command
   FullClose : BOOL;   // fully close the valve without ramp
   FullCloseSP : REAL;   // target value of the valve closing
   FullCloseResetTimer : TIMER;   // Timer to reset full close command
   ClosedStatusSP : REAL;   // Closed Status Setpoint
   ClosedStatus : BOOL;   // Closed Status
END_STRUCT
END_TYPE

TYPE Phases :   // Phase Control UDT
STRUCT
   Run : BOOL;   // Phase Run
   RunOSR : BOOL;   // Phase Run One-Shot
   Stop : BOOL;   // Phase Stop
   Hold : BOOL;   // Phase Hold
   Pause : BOOL;   // Phase Pause
   PauseOVR : BOOL;   // Pause Override
   Jump : BOOL;   // Phase Jump
   JumpPLC : BOOL;   // Phase Jump PLC
   Branch : BOOL;   // Branch Flag
   State : DINT;   // Phase State
   PendingStep : DINT;   // Pending Step Number
   JumpStep : DINT;   // Jump Step Number
   StartStep : DINT;   // Starting Step Number
   Crit1MetTime : DINT;   // Criteria 1 Met Timer
   NextStep : DINT;   // Next Step
   TotalSteps : DINT;   // Total Steps in Phase
   Label : DINT;   // Branch Label
   ActualStep : DINT;   // Actual Step
END_STRUCT
END_TYPE

TYPE PhaseTotalizer :   // Phase Totalizer UDT
STRUCT
   Enable : BOOL;   // Enable Totalizer
   PhaseEnable : BOOL;   // Enable Phase Totalizer
   StepEnable : BOOL;   // Enable Step Totalizer
   PauseEnable : BOOL;   // Enable Pause Totalizer
   UserEnable : BOOL;   // Enable User Totalizer
   ProcedureEnable : BOOL;   // Enable Procedure Totalizer
   PhaseReset : BOOL;   // Reset Phase Totalizer
   StepReset : BOOL;   // Reset Step Totalizer
   PauseReset : BOOL;   // Reset Pause Totalizer
   UserReset : BOOL;   // Reset User Totalizer
   PV : REAL;   // Totalizer Process Variable
   Phase : REAL;   // Phase Totalizer
   Step : REAL;   // Step Totalizer
   Pause : REAL;   // Pause Totalizer
   User : REAL;   // User Totalizer
   Procedure : REAL;   // Procedure Totalizer
   PVscale : REAL;   // PV Scaling
   PVsec : REAL;   // PV per second
   PVmin : REAL;   // PV Minimum Value
   Title : STRING10;   // Title to be displayed on status screen
   EGU : STRING10;   // EGU to display
   EnableCfg : BOOL;   // Set to one to use this totalizer
   SourceAddressCfg : INT;   // Enter analog Point # to be totalized
   SourceTypeCfg : BOOL;   // 0 For AnlogInput[] Source 1 For DerivedData.CVs Source
END_STRUCT
END_TYPE

TYPE PipeAnimation :   // Pipe Animation UDT
STRUCT
   PipeStat : BOOL[224];   // Pipe Animation Array
   PipeStatP1 : BOOL[224];   // Pipe Animation Array Line Pump 1
   PipeStatP2 : BOOL[224];   // Pipe Animation Array Line Pump 2
END_STRUCT
END_TYPE

TYPE Prompt :   // Prompt UDT
STRUCT
   Flag : BOOL;   // Flag
   PromptOK : BOOL;   // Type OK
   PromptYesNO : BOOL;   // Type Yes/No
   ResponseOK : BOOL;   // Input OK
   ResponseYes : BOOL;   // Input Yes
   ResponseNo : BOOL;   // Input No
   Pending : BOOL;   // Pending
   PromptONS : BOOL;   // One-Shot
   Step : DINT;   // Step Number
   Value : DINT;   // Value for PV+
END_STRUCT
END_TYPE

TYPE ScaleFiltering :   // Data for Scale Filtering
STRUCT
   CurrentFilter : INT;   // Type of filter used for Scale Filtering 0 = No Filtering 1 = Moving Average 2 = Exponential Linear Recursive
   Sample_Rate : DINT;   // Scale Filtering Sample Rate
   Timer : TIMER;   // Scale Filtering Timer
   WI001_Unfiltered : REAL;   // WI001 Unfiltered
   FeedBagVolume : REAL;   // Feed bag Volume based on WI001
   FeedBagVolume_Array : REAL[101];   // Array for Filter
   FeedBagVolume_MAVE : MOVING_AVERAGE;   // Feed Bag Volume Moving Average Filter structure
   FiltrateFlow : REAL;   // Filtrate Flow based on current filtrate volume
   FiltrateFlow_Array : REAL[101];   // Array for Filter
   FiltrateFlow_MAVE : MOVING_AVERAGE;   // Filtrate Flow Moving Average Filter structure
   FiltrateFlow_Mave_Timer : TIMER;   // Timer for MAVE Filter Flow
   FiltrateFlow_Mave_Sample_Rate : DINT;   // Filtrate Flow Sample Rate for MAVE
   FiltrateFlow_MaveFiltered : REAL;   // Filtrate Flow value filtered by MAVE
   FiltrateFlow_ExpConst : REAL;   // Constant for Exponential Filter
   FiltrateFlow_Exp_Timer : TIMER;   // Timer for Exponential Filter Flow
   FiltrateFlow_Exp_Sample_Rate : DINT;   // Filtrate Flow Sample Rate for Exp.
   FiltrateFlow_ExpFiltered : REAL;   // Filtrate Flow value filtered by Exp
   WI101_Unfiltered : REAL;   // WI101 Unfiltered
   FiltrateVolume101 : REAL;   // Filtrate Volume based on WI101
   FiltrateVolume101_Array : REAL[101];   // Array for Filter
   FiltrateVolume101_MAVE : MOVING_AVERAGE;   // Filtrate Volume 101 Moving Average Filter structure
   FiltrateVolume101_MaveFiltered : REAL;   // Filtrate Volume 101 value filtered by MAVE
   FiltrateVolume101_ExpConst : REAL;   // Constant for Exponential Filter
   FiltrateVolume101_ExpFiltered : REAL;   // Filtrate Volume 101 value filtered by Exp
   FiltrateVolume101_Filtered_Prev : REAL;   // Filtrate Volume 101 Filtered prev. Value
   Weight101_ExpFiltered : REAL;   // Filtrate Weight 101 filtered by Exp.
   Weight101_MaveFiltered : REAL;   // Filtrate Weight 101 filtered by MAVE
   WI102_Unfiltered : REAL;   // WI102 Unfiltered
   FiltrateVolume102 : REAL;   // Fitlrate Volume based on WI102
   FiltrateVolume102_Array : REAL[101];   // Array for Filter
   FiltrateVolume102_MAVE : MOVING_AVERAGE;   // Filtrate Volume 102 Moving Average Filter structure
   FiltrateVolume102_MaveFiltered : REAL;   // Filtrate Volume 102 value filtered by MAVE
   FiltrateVolume102_ExpConst : REAL;   // Constant for Exponential Filter
   FiltrateVolume102_ExpFiltered : REAL;   // Filtrate Volume 102 value filtered by Exp
   Weight102_ExpFiltered : REAL;   // Filtrate Weight 102 filtered by Exp.
   Weight102_MaveFiltered : REAL;   // Filtrate Weight 102 filtered by MAVE
   FiltrateVolume_ExpFiltered : REAL;   // Filtrate Volume Value filtered by Exp.
   FiltrateVolume_ExpFiltered_Prev : REAL;   // Filtrate Volume prev. Value filtered by Exp.
   FiltrateVolume_MaveFiltered : REAL;   // Filtrate Volume Value filtered by MAVE
   FiltrateVolume_MaveFiltered_Prev : REAL;   // Filtrate Volume prev. Value filtered by MAVE
END_STRUCT
END_TYPE

TYPE STRING10 :   // 10 Character String
STRUCT
   LEN : DINT;
   DATA : SINT[10];
END_STRUCT
END_TYPE

TYPE STRING240 :
STRUCT
   LEN : DINT;
   DATA : SINT[240];
END_STRUCT
END_TYPE

TYPE STRING25 :   // 25 Character String
STRUCT
   LEN : DINT;
   DATA : SINT[26];
END_STRUCT
END_TYPE

TYPE STRING4 :   // 4 Character String
STRUCT
   LEN : DINT;
   DATA : SINT[4];
END_STRUCT
END_TYPE

TYPE STRING5 :   // 5 Character String
STRUCT
   LEN : DINT;
   DATA : SINT[5];
END_STRUCT
END_TYPE

TYPE STRING50 :   // 50 Character String
STRUCT
   LEN : DINT;
   DATA : SINT[50];
END_STRUCT
END_TYPE

TYPE STRING6 :   // 6 Character String
STRUCT
   LEN : DINT;
   DATA : SINT[6];
END_STRUCT
END_TYPE

TYPE STRING80 :
STRUCT
   LEN : DINT;
   DATA : SINT[80];
END_STRUCT
END_TYPE

TYPE STRING90 :   // 90 Character String
STRUCT
   LEN : DINT;
   DATA : SINT[90];
END_STRUCT
END_TYPE

TYPE SysControl :   // System Control Mode UDT
STRUCT
   DefaultIn : BOOL;   // Set System in Default In
   DefaultOut : BOOL;   // Set System in Default Out
   DefaultTimer : TIMER;   // Set System in Default Timer
   AllAutoIn : BOOL;   // Set System in All Auto In
   AllAutoOut : BOOL;   // Set System in All Auto Out
   AllAutoTimer : TIMER;   // Set System in All Auto Timer
   Simulate : BOOL;   // Enable Simulation Mode
   Proc_Simulate : BOOL;   // Enable Process Simulation Mode
   Maintenance : BOOL;   // Enable Maintenance Mode
   DefaultStatus : BOOL;   // Default state status
   EnableSaveRestoreParam : BOOL;   // Enable save\restore parameters if condition are met
   UV_Auto_Zero_Cmd : BOOL;   // UV Auto Zero Command
   UV_Auto_Zero_Timer : TIMER;   // UV Auto Zero Timer
   Simulate_Options : BOOL;   // Allow Options simulation
END_STRUCT
END_TYPE

TYPE SystemType :   // System Type UDT
STRUCT
   StatusTimer : TIMER;   // Evaluate Status Value Delay Timer
   Value : INT;   // Current value of system type (0-none, 1-chrom, 2-TFF)
   MoldType : INT;   // Current Value of the Installed Mold (123=TF2S, 124=TF3S)
   HMI_Value : INT;   // Current value of system mold from HMI (123=TF2S, 124=TF3S)
   PreviousValue : INT;   // Previous selected value; used to determine if new selection is made
   EnableSystemType : BOOL[32];   // Enable System Types
   CopyConfigFromMoldType0 : BOOL[32];   // Copy configuration data from Mold Type 0 to all other Mold Types
   CopyConfigFromMoldType1 : BOOL[32];   // Copy configuration data from Mold Type 1 to all other Mold Types
   CopyConfigFromMoldType2 : BOOL[32];   // Copy configuration data from Mold Type 2 to all other Mold Types
   CopyConfigFromMoldType3 : BOOL[32];   // Copy configuration data from Mold Type 3 to all other Mold Types
   CopyConfigFromMoldType4 : BOOL[32];   // Copy configuration data from Mold Type 4 to all other Mold Types
   DisableStatusCheck : BOOL;   // Disable Status Check; Allows for manual setting of System Type
   Initialize : BOOL;   // Upon new system selection, Initialize bit is set for any system Initialization required for setting up new system type
   Error : BOOL;   // Error bit if unable to determine system type
   ChangeCS : BOOL;   // Change CS Action from HMI
   NewCS : BOOL;   // New CS detected
   CopyParametersActive : BOOL;   // Manually set bit before setting Copy Configuration Data
   NewSystem_Timer : TIMER;   // One-Minute System change Timer
END_STRUCT
END_TYPE

TYPE TankManagement :   // UDT to Manage Tank
STRUCT
   Config : TankRange;   // Tank Range Configuration Management
   WeightConfiguration : TankRangeParameters[4];   // Tank Weight Range Parameters Management
   LevelConfiguration : TankRangeParameters[4];   // Tank Level Range Parameters Management
   Feed_Bag_Tare : BOOL;   // Feed Bag Tare Command
   Feed_Bag_Tare_Timer : TIMER;   // Feed Bag Tare Timer for reset command
   Filtrate_Bag_Tare : BOOL;   // Filtrate Bag Tare Command
   Filtrate_Bag_Tare_Timer : TIMER;   // Filtrate Bag Tare Timer for reset command
END_STRUCT
END_TYPE

TYPE TankRange :   // Update Tank Range Scaling & Alarming
STRUCT
   TankSelected : DINT;   // Tank Selected (0-None, 1-TK50, 2-TK100, 3-TK250)
   TankSelectHMI : DINT;   // Tank Select HMI Use Only
   Option_Current : DINT;   // Tank Current Option
   Option_Prev : DINT;   // Tank Previous Option
   Option_Simulate : DINT;   // Tank Option Simulated
   TMR : TIMER;
   ONS : DINT;   // One Shots
   MismatchAlarm : BOOL;   // Detects if Tank Selected is different from the actual connected tank
   Accept : BOOL;   // Operator Accepts Tank Selection
   ForceUpdate : BOOL;   // Force Tank Selection Update even if Tank Selection is same as Connected Tank
   Update : BOOL;   // Tank Selection Update Required
   UpdateComplete : BOOL;   // Tank Selection Update Complete
   WTUseDefault : BOOL;   // Load Default Alarm SP values
   LTUseDefault : BOOL;   // Load Default Alarm SP values
   Simulate : BOOL;   // Simulate Tank Option (0-Off, 1-On)
   AlarmStatus : INT;   // Alarm Status ( 0 = No Alarm , 1 = Non Critical Alarm , 2 = Critical Alarm )
   LevelHMI : REAL;   // Tank Level scaled for Tank animation in HMI
END_STRUCT
END_TYPE

TYPE TankRangeParameters :   // Update Tank Range Scaling & Alarming
STRUCT
   Desc : STRING25;   // Description
   ScaledMin : REAL;   // Scaled Min
   ScaledMin_PRE : REAL;   // Scaled Min Previous
   ScaledMax : REAL;   // Scaled Max
   ScaledMax_PRE : REAL;   // Scaled Max Previous
   RangeMin : REAL;   // Range Min
   RangeMin_PRE : REAL;   // Range Min Previous
   RangeMax : REAL;   // Range Max
   RangeMax_PRE : REAL;   // Range Max Previous
   Alm_LOLO : REAL;   // LOLO Alarm SP
   Alm_LOLO_PRE : REAL;   // LOLO Alarm SP Previous
   Alm_LO : REAL;   // LO Alarm SP
   Alm_LO_PRE : REAL;   // LO Alarm SP Previous
   Alm_HI : REAL;   // HI Alarm SP
   Alm_HI_PRE : REAL;   // HI Alarm SP Previous
   Alm_HIHI : REAL;   // HIHI Alarm SP
   Alm_HIHI_PRE : REAL;   // HIHI Alarm SP Previous
   Alm_LOLOTMR : DINT;   // LOLO Alarm Timer Preset
   Alm_LOLOTMR_PRE : DINT;   // LOLO Alarm Timer Preset Previous
   Alm_LOTMR : DINT;   // LO Alarm Timer Preset
   Alm_LOTMR_PRE : DINT;   // LO Alarm Timer Preset Previous
   Alm_HITMR : DINT;   // HI Alarm Timer Preset
   Alm_HITMR_PRE : DINT;   // HI Alarm Timer Preset Previous
   Alm_HIHITMR : DINT;   // HIHI Alarm Timer Preset
   Alm_HIHITMR_PRE : DINT;   // HIHI Alarm Timer Preset Previous
   Alm_Override : BOOL;   // Alarm Override
END_STRUCT
END_TYPE

TYPE TimerControl :   // Timer Control UDT
STRUCT
   Tick : BOOL;   // 1 Second Tick
   TickMainTask : BOOL;   // 1 Second Tick to be used in MainTask
   NewTickMainTask : BOOL;   // Flag to triger the main task Tick
   ResetAll : BOOL;   // Reset All Timers/Totalizers
   ResetProcedure : BOOL;   // Reset Procedure Timers/Totalizers
   Save : DINT;   // Saved Timer Value
   Seconds : DINT;   // Master Seconds Value
   Colon : STRING4;   // Colon ":"
   ColonZero : STRING4;   // Colon with Zero ":0"
   Cycle : DINT;   // Compute Value each 25ms (cycle time of HighPriority Task)
END_STRUCT
END_TYPE

TYPE Timers :   // Timers UDT
STRUCT
   Enable : BOOL;   // Enable Timer
   Reset : BOOL;   // Reset Timer
   TotalSeconds : REAL;   // Total Seconds Value
   Hours : DINT;   // HH Integer Value
   Minutes : DINT;   // MM Integer Value
   Seconds : DINT;   // SS Integer Value
   sHours : STRING4;   // HH String Value
   sMinutes : STRING4;   // MM String Value
   sSeconds : STRING4;   // SS String Value
   HMS : STRING25;   // HH:MM:SS Value
   LastHMS : STRING25;   // HH:MM:SS Value
END_STRUCT
END_TYPE

TYPE Totalizers :   // Totalizers UDT
STRUCT
   Enable : BOOL;   // Enable Totalizer
   Reset : BOOL;   // Reset Phase Totalizer
   PV : REAL;   // Totalizer Process Variable
   Total : REAL;   // Phase Totalizer
   PVscale : REAL;   // PV Scaling
   PVsec : REAL;   // PV per second
   PVmin : REAL;   // PV Minimum Value
   Title : STRING10;   // Title to be displayed on status screen
   LastTotal : REAL;   // a copy of the total at the last reset
   ResetTimer : TIMER;   // Reset timer for event log
   ResetONS : BOOL;   // Reset one-shot
END_STRUCT
END_TYPE

TYPE UserAlarm :   // User Alarm UDT
STRUCT
   NonCritical1 : BOOL;   // Set the User Non Critical Alarm 1
   Critical1 : BOOL;   // Set the User Critical Alarm 1
   NonCritical2 : BOOL;   // Set the User Non Critical Alarm 2
   Critical2 : BOOL;   // Set the User Critical Alarm 2
   SetUserAlarm1ONS : BOOL;   // Set User Alarm 1 Oneshot
   SetUserAlarm2ONS : BOOL;   // Set User Alarm 2 Oneshot
END_STRUCT
END_TYPE

TYPE UserTotalizerManagement :   // User Totalizer Management UDT
STRUCT
   LogUserIn : BOOL;   // Log User Totalizer Value
   LogUserOut : BOOL;   // Log User Totalizer Value
   StartUser : BOOL;   // Start User Totalizer
   ResetUserIn : BOOL;   // Reset User Totalizer
   ResetUserOut : BOOL;   // Reset User Totalizer
   LogUserTimer : TIMER;   // Log User Totalizer Timer
   ResetUserTimer : TIMER;   // Reset User Totalizer Timer
END_STRUCT
END_TYPE

TYPE Valve :   // Valve UDT
STRUCT
   Tag : STRING5;   // Tag Name
   Desc : STRING25;   // Description
   Control : BOOL;   // Valve Control
   Auto : BOOL;   // Auto Command
   Manual : BOOL;   // Manual Command (Force)
   Mode : BOOL;   // Control Mode
   ZSOpen : BOOL;   // Open Limit Switch
   ZSClose : BOOL;   // Closed Limit Switch
   ZSOpenEnable : BOOL;   // Enable Open Limit Switch
   ZSCloseEnable : BOOL;   // Enable Closed Limit Switch
   OpenStatus : BOOL;   // Open/On Status
   CloseStatus : BOOL;   // Closed/Off Status
   ZSOverride : BOOL;   // Limit Switch Override
   Priority : BOOL;   // Alarm Priority 0=Low, 1=High
   PriorityCfg : BOOL;   // Set to 1 to allow user to set Priority and Enable
   Alarm : BOOL;   // Alarm
   AlarmAck : BOOL;   // Alarm Acknowledged
   FailState : BOOL;   // Fail State 0=Closed, 1=Open
   Ports : BOOL;   // Number of Ports 0=2 way, 1=3 way
   OpenONS : BOOL;   // Open One-Shot
   CloseONS : BOOL;   // Close One-Shot
   EnableCfg : BOOL;   // Set to 1 to activate this Tag
   StatusWord : DINT;   // Valve Status word for HMI
   Status : DINT;   // Valve Status for Audit Trail
   ZSOpenAddress : DINT;   // Open Limit Switch Input Address
   ZSCloseAddress : DINT;   // Closed Limit Switch Input Address
   OutputAddress : DINT;   // Valve Output Address
   AlarmTimer : TIMER;   // Alarm Timer
   AlarmTimerSP : DINT;   // Alarm Timer setpoint (sec)
   AutoCloseTimer : TIMER;   // Auto Close Timer
   AlarmONS : BOOL;   // One shot when alarm occurs
END_STRUCT
END_TYPE

TYPE ValveControl :   // Valve Control UDT
STRUCT
   NonCriticalFault : BOOL;   // Valve Non-Critical Fault
   NonCriticalFaultUnack : BOOL;   // Unacknowledged Valve Non-Critical Fault
   CriticalFault : BOOL;   // Valve Critical Fault
   CriticalFaultUnack : BOOL;   // Unacknowledged Valve Critical Fault
   ValveStatus1 : DINT;   // Valve Status (Valves 1-32)
   ValveStatus2 : DINT;   // Valve Status (Valves 33-64)
   ValveStatus3 : DINT;   // Valve Status (Valves 65-96)
   ValveStatus4 : DINT;   // Valve Status (Valves 97-128)
   Default1 : DINT;   // Default State (Valves 1-32)
   Default2 : DINT;   // Default State (Valves 33-64)
   Default3 : DINT;   // Default State (Valves 65-96)
   Default4 : DINT;   // Default State (Valves 97-128)
   MaxValveNum : DINT;   // Maximimum Valve Number
END_STRUCT
END_TYPE

TYPE XS_AlarmCond :   // AlarmCondition PrimingTimer or AlarmTime
STRUCT
   XS001_Enable : BOOL;   // Activate alarm
   XS001_Arm : BOOL;   // Select Priming Timer or Delay Timer
   XS001_PrimingTimer : DINT;   // Value of Priming Timer
   XS001_PrimingTimeSP : DINT;   // Priming Time set point (sec)
   XS001_Delaytimer : DINT;   // Value of Delay Timer
   XS001_AlarmTimeSP : DINT;   // Alarm Time set point (sec)
   XS002_Enable : BOOL;   // Activate alarm
   XS002_Arm : BOOL;   // Select Priming Timer or Delay Timer
   XS002_PrimingTimer : DINT;   // Value of Priming Timer
   XS002_PrimingTimeSP : DINT;   // Priming Time set point (sec)
   XS002_Delaytimer : DINT;   // Value of Delay Timer
   XS002_AlarmTimeSP : DINT;   // Alarm Time set point (sec)
END_STRUCT
END_TYPE

VAR_GLOBAL   (* controller tags *)
   ACQ002 : ALIAS FOR DigitalOutput[0];   // Emergency Stop Acknowledge
   AI101 : ALIAS FOR AnalogPoint[10];   // Filtrate Conductivity
   AI101_SIG : ALIAS FOR DigitalPoint[90];
   AI101Alarm : ALIAS FOR AlarmAnalog[10];   // Filtrate Conductivity Alarm
   AI102 : ALIAS FOR AnalogPoint[11];   // Filtrate UV
   AI102_SIG : ALIAS FOR DigitalPoint[91];
   AI102Alarm : ALIAS FOR AlarmAnalog[11];   // Filtrate UV Alarm
   AI103 : ALIAS FOR AnalogPoint[12];   // Filtrate UV
   AI103_SIG : ALIAS FOR DigitalPoint[92];
   AI103Alarm : ALIAS FOR AlarmAnalog[12];   // Filtrate UV Alarm
   AI104 : ALIAS FOR AnalogPoint[9];   // Filtrate pH
   AI104_SIG : ALIAS FOR DigitalPoint[105];
   AI104Alarm : ALIAS FOR AlarmAnalog[9];   // Filtrate pH Alarm
   AlarmAnalog : AlarmAnalog[50] := ([0].Override := 1, [0].LOLOAlarmONS := 1, [0].LOAlarmONS := 1, [0].HIAlarmONS := 1, [0].HIHIAlarmONS := 1, [0].HI := 1500.0, [0].HIHI := 1500.0, [0].LOLOTimer.PRE := 2000, [0].LOLOTimerSP := 2, [0].LOTimer.PRE := 2000, [0].LOTimerSP := 2, [0].HITimer.PRE := 2000, [0].HITimerSP := 2, [0].HIHITimer.PRE := 2000, [0].HIHITimerSP := 2, [1].Override := 1, [1].HI := 1000.0, [1].HIHI := 1000.0, [1].PV := -374.96228, [1].LOLOTimer.PRE := 2000, [1].LOLOTimerSP := 2, [1].LOTimer.PRE := 2000, [1].LOTimerSP := 2, [1].HITimer.PRE := 2000, [1].HITimerSP := 2, [1].HIHITimer.PRE := 2000, [1].HIHITimerSP := 2, [1].EnableCfg := 1, [2].Override := 1, [2].LOLODisable := 1, [2].LODisable := 1, [2].FeedPumpEnable := 1, [2].FeedPumpTag := 1, [2].HI := 19.8, [2].HIHI := 20.0, [2].LOLOTimer.PRE := 2000, [2].LOLOTimerSP := 2, [2].LOTimer.PRE := 2000, [2].LOTimerSP := 2, [2].HITimer.PRE := 2000, [2].HITimerSP := 2, [2].HIHITimer.PRE := 2000, [2].HIHITimerSP := 2, [2].EnableCfg := 1, [3].Override := 1, [3].HI := 100.0, [3].HIHI := 100.0, [3].PV := -3.499525, [3].LOLOTimer.PRE := 1000, [3].LOLOTimerSP := 2, [3].LOTimer.PRE := 5000, [3].LOTimerSP := 2, [3].HITimer.PRE := 5000, [3].HITimerSP := 2, [3].HIHITimer.PRE := 1000, [3].HIHITimerSP := 2, [4].Override := 1, [4].HI := 100.0, [4].HIHI := 100.0, [4].PV := -24.996607,
        [4].LOLOTimer.PRE := 1000, [4].LOLOTimerSP := 2, [4].LOTimer.PRE := 5000, [4].LOTimerSP := 2, [4].HITimer.PRE := 5000, [4].HITimerSP := 2, [4].HIHITimer.PRE := 1000, [4].HIHITimerSP := 2, [5].Override := 1, [5].LOLODisable := 1, [5].LODisable := 1, [5].HIHIEnable := 1, [5].FeedPumpEnable := 1, [5].FeedPumpTag := 1, [5].HI := 35.0, [5].HIHI := 38.0, [5].PV := 0.0066376748, [5].LOLOTimer.PRE := 2000, [5].LOLOTimerSP := 2, [5].LOTimer.PRE := 2000, [5].LOTimerSP := 2, [5].HITimer.PRE := 2000, [5].HITimerSP := 2, [5].HIHITimer.PRE := 2000, [5].HIHITimerSP := 2, [5].EnableCfg := 1, [6].Override := 1, [6].LOLODisable := 1, [6].LODisable := 1, [6].HIHIEnable := 1, [6].FeedPumpEnable := 1, [6].FeedPumpTag := 1, [6].HI := 40.0, [6].HIHI := 50.0, [6].PV := -0.21904327, [6].LOLOTimer.PRE := 2000, [6].LOLOTimerSP := 2, [6].LOTimer.PRE := 2000, [6].LOTimerSP := 2, [6].HITimer.PRE := 2000, [6].HITimerSP := 2, [6].HIHITimer.PRE := 2000, [6].HIHITimerSP := 2, [6].EnableCfg := 1, [7].Override := 1, [7].LOLODisable := 1, [7].LODisable := 1, [7].HIHIEnable := 1, [7].FeedPumpEnable := 1, [7].FeedPumpTag := 1, [7].HI := 18.0, [7].HIHI := 20.0, [7].PV := -0.22568095, [7].LOLOTimer.PRE := 2000, [7].LOLOTimerSP := 2, [7].LOTimer.PRE := 2000, [7].LOTimerSP := 2, [7].HITimer.PRE := 2000, [7].HITimerSP := 2, [7].HIHITimer.PRE := 2000,
        [7].HIHITimerSP := 2, [7].EnableCfg := 1, [8].Override := 1, [8].LOLODisable := 1, [8].LODisable := 1, [8].HIHIEnable := 1, [8].TransferPumpEnable := 1, [8].TransferPumpTag := 2, [8].HI := 40.0, [8].HIHI := 50.0, [8].PV := 0.2920577, [8].LOLOTimer.PRE := 2000, [8].LOLOTimerSP := 2, [8].LOTimer.PRE := 2000, [8].LOTimerSP := 2, [8].HITimer.PRE := 2000, [8].HITimerSP := 2, [8].HIHITimer.PRE := 2000, [8].HIHITimerSP := 2, [8].EnableCfg := 1, [9].Override := 1, [9].HI := 14.0, [9].HIHI := 14.0, [9].PV := -1.4998856, [9].LOLOTimer.PRE := 2000, [9].LOLOTimerSP := 2, [9].LOTimer.PRE := 2000, [9].LOTimerSP := 2, [9].HITimer.PRE := 2000, [9].HITimerSP := 2, [9].HIHITimer.PRE := 2000, [9].HIHITimerSP := 2, [10].Override := 1, [10].HI := 180.0, [10].HIHI := 200.0, [10].PV := 0.030518044, [10].LOLOTimer.PRE := 2000, [10].LOLOTimerSP := 2, [10].LOTimer.PRE := 2000, [10].LOTimerSP := 2, [10].HITimer.PRE := 2000, [10].HITimerSP := 2, [10].HIHITimer.PRE := 2000, [10].HIHITimerSP := 2, [10].EnableCfg := 1, [11].Override := 1, [11].HI := 0.5, [11].HIHI := 0.8, [11].PV := 0.09529259, [11].LOLOTimer.PRE := 2000, [11].LOLOTimerSP := 2, [11].LOTimer.PRE := 2000, [11].LOTimerSP := 2, [11].HITimer.PRE := 2000, [11].HITimerSP := 2, [11].HIHITimer.PRE := 2000, [11].HIHITimerSP := 2, [11].EnableCfg := 1, [12].Override := 1, [12].HI := 0.5,
        [12].HIHI := 0.8, [12].PV := 0.030975815, [12].LOLOTimer.PRE := 2000, [12].LOLOTimerSP := 2, [12].LOTimer.PRE := 2000, [12].LOTimerSP := 2, [12].HITimer.PRE := 2000, [12].HITimerSP := 2, [12].HIHITimer.PRE := 2000, [12].HIHITimerSP := 2, [12].EnableCfg := 1, [13].Override := 1, [13].HI := 45.0, [13].HIHI := 55.0, [13].PV := 20.54265, [13].LOLOTimer.PRE := 2000, [13].LOLOTimerSP := 2, [13].LOTimer.PRE := 2000, [13].LOTimerSP := 2, [13].HITimer.PRE := 2000, [13].HITimerSP := 2, [13].HIHITimer.PRE := 2000, [13].HIHITimerSP := 2, [13].EnableCfg := 1, [14].Override := 1, [14].HI := 100.0, [14].HIHI := 100.0, [14].LOLOTimerSP := 2, [14].LOTimerSP := 2, [14].HITimerSP := 2, [14].HIHITimerSP := 2, [15].Override := 1, [15].LOLODisable := 1, [15].LODisable := 1, [15].FeedPumpEnable := 1, [15].FeedPumpTag := 1, [15].HI := 230.0, [15].HIHI := 240.0, [15].EnableCfg := 1, [16].Override := 1, [16].PV := -0.4999322, [16].LOLOTimerSP := 2, [16].LOTimerSP := 2, [16].HITimerSP := 2, [16].HIHITimerSP := 2, [17].Override := 1, [17].FeedPumpEnable := 1, [17].TransferPumpEnable := 1, [17].FeedPumpTag := 1, [17].TransferPumpTag := 2, [17].PV := -2.499796, [17].LOLOTimerSP := 2, [17].LOTimerSP := 2, [17].HITimerSP := 2, [17].HIHITimerSP := 2, [18].Override := 1, [18].PV := -2.499796, [18].LOLOTimerSP := 2, [18].LOTimerSP := 2, [18].HITimerSP := 2,
        [18].HIHITimerSP := 2, [19].Override := 1, [19].PV := -2.499796, [19].LOLOTimerSP := 2, [19].LOTimerSP := 2, [19].HITimerSP := 2, [19].HIHITimerSP := 2, [20].Override := 1, [20].PV := 100.0, [20].LOLOTimerSP := 2, [20].LOTimerSP := 2, [20].HITimer.EN := 1, [20].HITimer.DN := 1, [20].HITimerSP := 2, [20].HIHITimer.EN := 1, [20].HIHITimer.DN := 1, [20].HIHITimerSP := 2, [21].Override := 1, [21].LOLOTimerSP := 2, [21].LOTimerSP := 2, [21].HITimerSP := 2, [21].HIHITimerSP := 2, [22].Override := 1, [22].PV := 0.5047684, [23].Override := 1, [23].PV := 0.1161975, [24].Override := 1, [24].PV := 0.16, [25].Override := 1, [25].PV := -0.3333333, [26].Override := 1, [26].PV := 63.88032, [27].Override := 1, [27].PV := -37.40687, [28].Override := 1, [28].HI := 100.0, [28].HIHI := 100.0, [28].PV := 22.8542, [28].LOLOTimer.PRE := 2000, [28].LOLOTimerSP := 2, [28].LOTimer.PRE := 2000, [28].LOTimerSP := 2, [28].HITimer.PRE := 2000, [28].HITimerSP := 2, [28].HIHITimer.PRE := 2000, [28].HIHITimerSP := 2, [29].Override := 1, [29].HI := 100.0, [29].HIHI := 100.0, [29].PV := 21.877623, [29].LOLOTimer.PRE := 2000, [29].LOLOTimerSP := 2, [29].LOTimer.PRE := 2000, [29].LOTimerSP := 2, [29].HITimer.PRE := 2000, [29].HITimerSP := 2, [29].HIHITimer.PRE := 2000, [29].HIHITimerSP := 2, [30].Override := 1, [30].HI := 100.0,
        [30].HIHI := 100.0, [30].PV := 21.877623, [30].LOLOTimer.PRE := 2000, [30].LOLOTimerSP := 2, [30].LOTimer.PRE := 2000, [30].LOTimerSP := 2, [30].HITimer.PRE := 2000, [30].HITimerSP := 2, [30].HIHITimer.PRE := 2000, [30].HIHITimerSP := 2, [31].Override := 1, [31].HI := 100.0, [31].HIHI := 100.0, [31].PV := 21.877623, [31].LOLOTimer.PRE := 2000, [31].LOLOTimerSP := 2, [31].LOTimer.PRE := 2000, [31].LOTimerSP := 2, [31].HITimer.PRE := 2000, [31].HITimerSP := 2, [31].HIHITimer.PRE := 2000, [31].HIHITimerSP := 2, [32].Override := 1, [32].PV := 0.1837702, [33].Override := 1, [33].PV := -0.6615715, [34].Override := 1, [34].PV := 0.6615715, [35].Override := 1, [35].PV := 222.0, [36].Override := 1, [37].Override := 1, [37].PV := -0.03181506, [38].Override := 1, [39].Override := 1, [40].Override := 1, [40].LOLODisable := 1, [40].LODisable := 1, [40].FeedPumpEnable := 1, [40].FeedPumpTag := 1, [40].HI := 75.0, [40].HIHI := 87.0, [40].PV := 0.30865186, [40].LOLOTimer.PRE := 2000, [40].LOLOTimerSP := 2, [40].LOTimer.PRE := 2000, [40].LOTimerSP := 2, [40].HITimer.PRE := 2000, [40].HITimerSP := 2, [40].HIHITimer.PRE := 2000, [40].HIHITimerSP := 2, [40].EnableCfg := 1, [41].Override := 1, [41].LOLODisable := 1, [41].LODisable := 1, [41].FeedPumpEnable := 1, [41].FeedPumpTag := 1, [41].HI := 75.0, [41].HIHI := 87.0, [41].PV := 0.087949194,
        [41].LOLOTimer.PRE := 2000, [41].LOLOTimerSP := 2, [41].LOTimer.PRE := 2000, [41].LOTimerSP := 2, [41].HITimer.PRE := 2000, [41].HITimerSP := 2, [41].HIHITimer.PRE := 2000, [41].HIHITimerSP := 2, [41].EnableCfg := 1, [42].Override := 1, [42].LOLODisable := 1, [42].LODisable := 1, [42].FeedPumpEnable := 1, [42].FeedPumpTag := 1, [42].HI := 40.0, [42].HIHI := 44.0, [42].LOLOTimer.PRE := 2000, [42].LOLOTimerSP := 2, [42].LOTimer.PRE := 2000, [42].LOTimerSP := 2, [42].HITimer.PRE := 2000, [42].HITimerSP := 2, [42].HIHITimer.PRE := 2000, [42].HIHITimerSP := 2, [42].EnableCfg := 1, [43].Override := 1, [43].LOLODisable := 1, [43].LODisable := 1, [43].TransferPumpEnable := 1, [43].TransferPumpTag := 2, [43].HI := 20.0, [43].HIHI := 22.0, [43].LOLOTimer.PRE := 2000, [43].LOLOTimerSP := 2, [43].LOTimer.PRE := 2000, [43].LOTimerSP := 2, [43].HITimer.PRE := 2000, [43].HITimerSP := 2, [43].HIHITimer.PRE := 2000, [43].HIHITimerSP := 2, [43].EnableCfg := 1, [44].Override := 1, [44].LOLODisable := 1, [44].LODisable := 1, [44].FeedPumpEnable := 1, [44].FeedPumpTag := 1, [44].HI := 190.0, [44].HIHI := 200.0, [44].EnableCfg := 1, [45].Override := 1, [45].HI := 999.0, [45].HIHI := 999.0, [45].LOLOTimerSP := 2, [45].LOTimerSP := 2, [45].HITimerSP := 2, [45].HIHITimerSP := 2, [46].Override := 1, [46].HI := 999.0, [46].HIHI := 999.0, [46].LOLOTimerSP := 2,
        [46].LOTimerSP := 2, [46].HITimerSP := 2, [46].HIHITimerSP := 2, [47].Override := 1, [48].Override := 1, [49].Override := 1);   // Analog Alarm Array
        [10]   // FI001Alarm
        [11]   // PI001Alarm
        [12]   // FI002Alarm
        [1]   // AI201BAlarm
        [2]   // AI201AAlarm
        [13]   // PI002Alarm
        [17]   // FI003Alarm
        [40]   // FI003Alarm
        [3]   // AI202Alarm
        [4]   // TI201Alarm
        [41]   // LV003Alarm
        [42]   // LV001Alarm
        [43]   // LV002Alarm
        [5]   // AI203Alarm
        [6]   // AI204Alarm
        [7]   // AI102Alarm
        [8]   // AI103Alarm
        [9]   // PI003Alarm
   AlarmAnalog_Storage : AlarmAnalog[6,50] := ([0,0].LOLOAlarmONS := 1, [0,0].LOAlarmONS := 1, [0,0].HIAlarmONS := 1, [0,0].HIHIAlarmONS := 1, [0,0].HI := 100.0, [0,0].HIHI := 100.0, [0,0].PV := -2.4997964, [0,0].LOLOTimer.PRE := 2000, [0,0].LOLOTimerSP := 2, [0,0].LOTimer.PRE := 2000, [0,0].LOTimerSP := 2, [0,0].HITimer.PRE := 2000, [0,0].HITimerSP := 2, [0,0].HIHITimer.PRE := 2000, [0,0].HIHITimerSP := 2, [0,1].HI := 50.0, [0,1].HIHI := 50.0, [0,1].PV := -12.498303, [0,1].LOLOTimer.PRE := 2000, [0,1].LOLOTimerSP := 2, [0,1].LOTimer.PRE := 2000, [0,1].LOTimerSP := 2, [0,1].HITimer.PRE := 2000, [0,1].HITimerSP := 2, [0,1].HIHITimer.PRE := 2000, [0,1].HIHITimerSP := 2, [0,1].EnableCfg := 1, [0,2].HI := 100.0, [0,2].HIHI := 100.0, [0,2].PV := -24.996607, [0,2].LOLOTimer.PRE := 2000, [0,2].LOLOTimerSP := 2, [0,2].LOTimer.PRE := 2000, [0,2].LOTimerSP := 2, [0,2].HITimer.PRE := 2000, [0,2].HITimerSP := 2, [0,2].HIHITimer.PRE := 2000, [0,2].HIHITimerSP := 2, [0,2].EnableCfg := 1, [0,3].HI := 14.0, [0,3].HIHI := 14.0, [0,3].PV := -3.499525, [0,3].LOLOTimer.PRE := 1000, [0,3].LOLOTimerSP := 1, [0,3].LOTimer.PRE := 5000, [0,3].LOTimerSP := 5, [0,3].HITimer.PRE := 5000, [0,3].HITimerSP := 5, [0,3].HIHITimer.PRE := 1000, [0,3].HIHITimerSP := 1, [0,3].EnableCfg := 1, [0,4].HI := 100.0, [0,4].HIHI := 100.0, [0,4].PV := -24.996607, [0,4].LOLOTimer.PRE := 1000, [0,4].LOLOTimerSP := 1, [0,4].LOTimer.PRE := 5000, [0,4].LOTimerSP := 5, [0,4].HITimer.PRE := 5000, [0,4].HITimerSP := 5,
        [0,4].HIHITimer.PRE := 1000, [0,4].HIHITimerSP := 1, [0,4].EnableCfg := 1, [0,5].HI := 2.0, [0,5].HIHI := 2.0, [0,5].PV := -0.49993217, [0,5].LOLOTimer.PRE := 2000, [0,5].LOLOTimerSP := 2, [0,5].LOTimer.PRE := 2000, [0,5].LOTimerSP := 2, [0,5].HITimer.PRE := 2000, [0,5].HITimerSP := 2, [0,5].HIHITimer.PRE := 2000, [0,5].HIHITimerSP := 2, [0,5].EnableCfg := 1, [0,6].HI := 2.0, [0,6].HIHI := 2.0, [0,6].PV := -0.49993217, [0,6].LOLOTimer.PRE := 2000, [0,6].LOLOTimerSP := 2, [0,6].LOTimer.PRE := 2000, [0,6].LOTimerSP := 2, [0,6].HITimer.PRE := 2000, [0,6].HITimerSP := 2, [0,6].HIHITimer.PRE := 2000, [0,6].HIHITimerSP := 2, [0,6].EnableCfg := 1, [0,7].HI := 100.0, [0,7].HIHI := 100.0, [0,7].PV := -24.996607, [0,7].LOLOTimer.PRE := 2000, [0,7].LOLOTimerSP := 2, [0,7].LOTimer.PRE := 2000, [0,7].LOTimerSP := 2, [0,7].HITimer.PRE := 2000, [0,7].HITimerSP := 2, [0,7].HIHITimer.PRE := 2000, [0,7].HIHITimerSP := 2, [0,7].EnableCfg := 1, [0,8].HI := 14.0, [0,8].HIHI := 14.0, [0,8].PV := -3.499525, [0,8].LOLOTimer.PRE := 1000, [0,8].LOLOTimerSP := 1, [0,8].LOTimer.PRE := 5000, [0,8].LOTimerSP := 5, [0,8].HITimer.PRE := 5000, [0,8].HITimerSP := 5, [0,8].HIHITimer.PRE := 1000, [0,8].HIHITimerSP := 1, [0,8].EnableCfg := 1, [0,9].LOLODisable := 1, [0,9].LODisable := 1, [0,9].FeedPumpEnable := 1, [0,9].TransferPumpEnable := 1, [0,9].FeedPumpTag := 1, [0,9].TransferPumpTag := 2, [0,9].HI := 6.0, [0,9].HIHI := 6.0, [0,9].PV := -1.4998856,
        [0,9].LOLOTimer.PRE := 2000, [0,9].LOLOTimerSP := 2, [0,9].LOTimer.PRE := 2000, [0,9].LOTimerSP := 2, [0,9].HITimer.PRE := 2000, [0,9].HITimerSP := 2, [0,9].HIHITimer.PRE := 2000, [0,9].HIHITimerSP := 2, [0,9].EnableCfg := 1, [0,10].LOLODisable := 1, [0,10].LODisable := 1, [0,10].FeedPumpEnable := 1, [0,10].FeedPumpTag := 1, [0,10].HI := 22.0, [0,10].HIHI := 22.0, [0,10].LOLOTimer.PRE := 2000, [0,10].LOLOTimerSP := 2, [0,10].LOTimer.PRE := 2000, [0,10].LOTimerSP := 2, [0,10].HITimer.PRE := 2000, [0,10].HITimerSP := 2, [0,10].HIHITimer.PRE := 2000, [0,10].HIHITimerSP := 2, [0,10].EnableCfg := 1, [0,11].LOLODisable := 1, [0,11].LODisable := 1, [0,11].FeedPumpEnable := 1, [0,11].FeedPumpTag := 1, [0,11].HI := 6.0, [0,11].HIHI := 6.0, [0,11].PV := -1.4998856, [0,11].LOLOTimer.PRE := 2000, [0,11].LOLOTimerSP := 2, [0,11].LOTimer.PRE := 2000, [0,11].LOTimerSP := 2, [0,11].HITimer.PRE := 2000, [0,11].HITimerSP := 2, [0,11].HIHITimer.PRE := 2000, [0,11].HIHITimerSP := 2, [0,11].EnableCfg := 1, [0,12].LOLODisable := 1, [0,12].LODisable := 1, [0,12].TransferPumpEnable := 1, [0,12].TransferPumpTag := 2, [0,12].HI := 22.0, [0,12].HIHI := 22.0, [0,12].LOLOTimer.PRE := 2000, [0,12].LOLOTimerSP := 2, [0,12].LOTimer.PRE := 2000, [0,12].LOTimerSP := 2, [0,12].HITimer.PRE := 2000, [0,12].HITimerSP := 2, [0,12].HIHITimer.PRE := 2000, [0,12].HIHITimerSP := 2, [0,12].EnableCfg := 1, [0,13].LOLODisable := 1, [0,13].LODisable := 1, [0,13].TransferPumpEnable := 1, [0,13].TransferPumpTag := 2, [0,13].HI := 6.0,
        [0,13].HIHI := 6.0, [0,13].PV := -1.4998856, [0,13].LOLOTimer.PRE := 2000, [0,13].LOLOTimerSP := 2, [0,13].LOTimer.PRE := 2000, [0,13].LOTimerSP := 2, [0,13].HITimer.PRE := 2000, [0,13].HITimerSP := 2, [0,13].HIHITimer.PRE := 2000, [0,13].HIHITimerSP := 2, [0,13].EnableCfg := 1, [0,14].Override := 1, [0,14].HI := 14.0, [0,14].HIHI := 14.0, [0,14].LOLOTimer.PRE := 1000, [0,14].LOLOTimerSP := 1, [0,14].LOTimer.PRE := 5000, [0,14].LOTimerSP := 5, [0,14].HITimer.PRE := 5000, [0,14].HITimerSP := 5, [0,14].HIHITimer.PRE := 1000, [0,14].HIHITimerSP := 1, [0,15].Override := 1, [0,15].HI := 2.0, [0,15].HIHI := 2.0, [0,15].PV := -0.49993217, [0,15].LOLOTimer.PRE := 2000, [0,15].LOLOTimerSP := 2, [0,15].LOTimer.PRE := 2000, [0,15].LOTimerSP := 2, [0,15].HITimer.PRE := 2000, [0,15].HITimerSP := 2, [0,15].HIHITimer.PRE := 2000, [0,15].HIHITimerSP := 2, [0,16].Override := 1, [0,16].HI := 2.0, [0,16].HIHI := 2.0, [0,16].PV := -0.49993217, [0,16].LOLOTimer.PRE := 2000, [0,16].LOLOTimerSP := 2, [0,16].LOTimer.PRE := 2000, [0,16].LOTimerSP := 2, [0,16].HITimer.PRE := 2000, [0,16].HITimerSP := 2, [0,16].HIHITimer.PRE := 2000, [0,16].HIHITimerSP := 2, [0,17].Override := 1, [0,17].FeedPumpEnable := 1, [0,17].TransferPumpEnable := 1, [0,17].FeedPumpTag := 1, [0,17].TransferPumpTag := 2, [0,17].LOLO := -1.0, [0,17].LO := -1.0, [0,17].HI := 5.0, [0,17].HIHI := 5.0, [0,17].PV := -2.4997964, [0,17].LOLOTimer.PRE := 2000, [0,17].LOLOTimerSP := 2, [0,17].LOTimer.PRE := 2000, [0,17].LOTimerSP := 2,
        [0,17].HITimer.PRE := 2000, [0,17].HITimerSP := 2, [0,17].HIHITimer.PRE := 2000, [0,17].HIHITimerSP := 2, [0,18].Override := 1, [0,18].FeedPumpEnable := 1, [0,18].FeedPumpTag := 1, [0,18].LOLO := -1.0, [0,18].LO := -1.0, [0,18].HI := 5.0, [0,18].HIHI := 5.0, [0,18].PV := -2.4997964, [0,18].LOLOTimer.PRE := 2000, [0,18].LOLOTimerSP := 2, [0,18].LOTimer.PRE := 2000, [0,18].LOTimerSP := 2, [0,18].HITimer.PRE := 2000, [0,18].HITimerSP := 2, [0,18].HIHITimer.PRE := 2000, [0,18].HIHITimerSP := 2, [0,19].Override := 1, [0,19].TransferPumpEnable := 1, [0,19].TransferPumpTag := 2, [0,19].LOLO := -1.0, [0,19].LO := -1.0, [0,19].HI := 5.0, [0,19].HIHI := 5.0, [0,19].PV := -2.4997964, [0,19].LOLOTimer.PRE := 2000, [0,19].LOLOTimerSP := 2, [0,19].LOTimer.PRE := 2000, [0,19].LOTimerSP := 2, [0,19].HITimer.PRE := 2000, [0,19].HITimerSP := 2, [0,19].HIHITimer.PRE := 2000, [0,19].HIHITimerSP := 2, [0,20].Override := 1, [0,20].HI := 100.0, [0,20].HIHI := 100.0, [0,20].PV := 100.0, [0,20].LOLOTimerSP := 2, [0,20].LOTimerSP := 2, [0,20].HITimer.EN := 1, [0,20].HITimer.DN := 1, [0,20].HITimerSP := 2, [0,20].HIHITimer.EN := 1, [0,20].HIHITimer.DN := 1, [0,20].HIHITimerSP := 2, [0,21].Override := 1, [0,21].HI := 100.0, [0,21].HIHI := 100.0, [0,21].LOLOTimerSP := 2, [0,21].LOTimerSP := 2, [0,21].HITimerSP := 2, [0,21].HIHITimerSP := 2, [0,22].Override := 1, [0,22].PV := 0.50476843, [0,23].Override := 1, [0,23].PV := 0.11619745, [0,24].Override := 1,
        [0,24].PV := 0.16, [0,25].Override := 1, [0,25].PV := -0.3333333, [0,26].Override := 1, [0,26].PV := 63.88032, [0,27].Override := 1, [0,27].PV := -37.40687, [0,28].HI := 100.0, [0,28].HIHI := 100.0, [0,28].PV := -24.998093, [0,28].LOLOTimer.PRE := 2000, [0,28].LOLOTimerSP := 2, [0,28].LOTimer.PRE := 2000, [0,28].LOTimerSP := 2, [0,28].HITimer.PRE := 2000, [0,28].HITimerSP := 2, [0,28].HIHITimer.PRE := 2000, [0,28].HIHITimerSP := 2, [0,28].EnableCfg := 1, [0,29].HI := 100.0, [0,29].HIHI := 100.0, [0,29].PV := -24.998093, [0,29].LOLOTimer.PRE := 2000, [0,29].LOLOTimerSP := 2, [0,29].LOTimer.PRE := 2000, [0,29].LOTimerSP := 2, [0,29].HITimer.PRE := 2000, [0,29].HITimerSP := 2, [0,29].HIHITimer.PRE := 2000, [0,29].HIHITimerSP := 2, [0,29].EnableCfg := 1, [0,30].HI := 100.0, [0,30].HIHI := 100.0, [0,30].PV := -24.811169, [0,30].LOLOTimer.PRE := 2000, [0,30].LOLOTimerSP := 2, [0,30].LOTimer.PRE := 2000, [0,30].LOTimerSP := 2, [0,30].HITimer.PRE := 2000, [0,30].HITimerSP := 2, [0,30].HIHITimer.PRE := 2000, [0,30].HIHITimerSP := 2, [0,30].EnableCfg := 1, [0,31].HI := 100.0, [0,31].HIHI := 100.0, [0,31].PV := -24.814985, [0,31].LOLOTimer.PRE := 2000, [0,31].LOLOTimerSP := 2, [0,31].LOTimer.PRE := 2000, [0,31].LOTimerSP := 2, [0,31].HITimer.PRE := 2000, [0,31].HITimerSP := 2, [0,31].HIHITimer.PRE := 2000, [0,31].HIHITimerSP := 2, [0,31].EnableCfg := 1, [0,32].Override := 1, [0,32].PV := 0.1837702, [0,33].Override := 1, [0,33].PV := -0.6615715, [0,34].Override := 1,
        [0,34].PV := 0.6615715, [0,35].Override := 1, [0,35].PV := 222.0, [0,36].Override := 1, [0,37].Override := 1, [0,37].PV := -0.03181506, [0,38].Override := 1, [0,39].Override := 1, [0,40].LOLODisable := 1, [0,40].LODisable := 1, [0,40].FeedPumpEnable := 1, [0,40].TransferPumpEnable := 1, [0,40].FeedPumpTag := 1, [0,40].TransferPumpTag := 2, [0,40].HI := 44.0, [0,40].HIHI := 44.0, [0,40].LOLOTimer.PRE := 2000, [0,40].LOLOTimerSP := 2, [0,40].LOTimer.PRE := 2000, [0,40].LOTimerSP := 2, [0,40].HITimer.PRE := 2000, [0,40].HITimerSP := 2, [0,40].HIHITimer.PRE := 2000, [0,40].HIHITimerSP := 2, [0,40].EnableCfg := 1, [0,41].LOLODisable := 1, [0,41].LODisable := 1, [0,41].FeedPumpEnable := 1, [0,41].TransferPumpEnable := 1, [0,41].FeedPumpTag := 1, [0,41].TransferPumpTag := 2, [0,41].HI := 9999.0, [0,41].HIHI := 9999.0, [0,41].LOLOTimer.PRE := 2000, [0,41].LOLOTimerSP := 2, [0,41].LOTimer.PRE := 2000, [0,41].LOTimerSP := 2, [0,41].HITimer.PRE := 2000, [0,41].HITimerSP := 2, [0,41].HIHITimer.PRE := 2000, [0,41].HIHITimerSP := 2, [0,41].EnableCfg := 1, [0,42].LOLODisable := 1, [0,42].LODisable := 1, [0,42].FeedPumpEnable := 1, [0,42].FeedPumpTag := 1, [0,42].HI := 9999.0, [0,42].HIHI := 9999.0, [0,42].LOLOTimer.PRE := 2000, [0,42].LOLOTimerSP := 2, [0,42].LOTimer.PRE := 2000, [0,42].LOTimerSP := 2, [0,42].HITimer.PRE := 2000, [0,42].HITimerSP := 2, [0,42].HIHITimer.PRE := 2000, [0,42].HIHITimerSP := 2, [0,42].EnableCfg := 1, [0,43].LOLODisable := 1, [0,43].LODisable := 1, [0,43].TransferPumpEnable := 1,
        [0,43].TransferPumpTag := 2, [0,43].HI := 9999.0, [0,43].HIHI := 9999.0, [0,43].LOLOTimer.PRE := 2000, [0,43].LOLOTimerSP := 2, [0,43].LOTimer.PRE := 2000, [0,43].LOTimerSP := 2, [0,43].HITimer.PRE := 2000, [0,43].HITimerSP := 2, [0,43].HIHITimer.PRE := 2000, [0,43].HIHITimerSP := 2, [0,43].EnableCfg := 1, [0,44].Override := 1, [0,44].HI := 99999.0, [0,44].HIHI := 99999.0, [0,44].LOLOTimerSP := 2, [0,44].LOTimerSP := 2, [0,44].HITimerSP := 2, [0,44].HIHITimerSP := 2, [0,45].Override := 1, [0,45].Disable := 1, [0,45].FeedPumpEnable := 1, [0,45].TransferPumpEnable := 1, [0,45].FeedPumpTag := 1, [0,45].TransferPumpTag := 2, [0,45].LOLO := -1.0, [0,45].LO := -1.0, [0,45].HI := 5.0, [0,45].HIHI := 5.0, [0,45].LOLOTimer.PRE := 2000, [0,45].LOLOTimerSP := 2, [0,45].LOTimer.PRE := 2000, [0,45].LOTimerSP := 2, [0,45].HITimer.PRE := 2000, [0,45].HITimerSP := 2, [0,45].HIHITimer.PRE := 2000, [0,45].HIHITimerSP := 2, [0,46].Override := 1, [0,47].Override := 1, [0,48].Override := 1, [0,49].Override := 1, [1,0].HI := 600.0, [1,0].HIHI := 600.0, [1,0].LOLOTimer.PRE := 2000, [1,0].LOLOTimerSP := 2, [1,0].LOTimer.PRE := 2000, [1,0].LOTimerSP := 2, [1,0].HITimer.PRE := 2000, [1,0].HITimerSP := 2, [1,0].HIHITimer.PRE := 2000, [1,0].HIHITimerSP := 2, [1,0].EnableCfg := 1, [1,1].Override := 1, [1,1].HI := 1000.0, [1,1].HIHI := 1000.0, [1,1].LOLOTimer.PRE := 2000, [1,1].LOLOTimerSP := 2, [1,1].LOTimer.PRE := 2000, [1,1].LOTimerSP := 2, [1,1].HITimer.PRE := 2000,
        [1,1].HITimerSP := 2, [1,1].HIHITimer.PRE := 2000, [1,1].HIHITimerSP := 2, [1,2].LOLODisable := 1, [1,2].LODisable := 1, [1,2].FeedPumpEnable := 1, [1,2].FeedPumpTag := 1, [1,2].HI := 15.0, [1,2].HIHI := 15.0, [1,2].PV := 0.01201648, [1,2].LOLOTimer.PRE := 2000, [1,2].LOLOTimerSP := 2, [1,2].LOTimer.PRE := 2000, [1,2].LOTimerSP := 2, [1,2].HITimer.PRE := 2000, [1,2].HITimerSP := 2, [1,2].HIHITimer.PRE := 2000, [1,2].HIHITimerSP := 2, [1,2].EnableCfg := 1, [1,3].Override := 1, [1,3].HI := 100.0, [1,3].HIHI := 100.0, [1,3].LOLOTimer.PRE := 1000, [1,3].LOLOTimerSP := 2, [1,3].LOTimer.PRE := 5000, [1,3].LOTimerSP := 2, [1,3].HITimer.PRE := 5000, [1,3].HITimerSP := 2, [1,3].HIHITimer.PRE := 1000, [1,3].HIHITimerSP := 2, [1,4].Override := 1, [1,4].HI := 100.0, [1,4].HIHI := 100.0, [1,4].LOLOTimer.PRE := 1000, [1,4].LOLOTimerSP := 2, [1,4].LOTimer.PRE := 5000, [1,4].LOTimerSP := 2, [1,4].HITimer.PRE := 5000, [1,4].HITimerSP := 2, [1,4].HIHITimer.PRE := 1000, [1,4].HIHITimerSP := 2, [1,5].LOLODisable := 1, [1,5].LODisable := 1, [1,5].HIHIEnable := 1, [1,5].FeedPumpEnable := 1, [1,5].FeedPumpTag := 1, [1,5].HI := 6.0, [1,5].HIHI := 6.0, [1,5].PV := -0.010986496, [1,5].LOLOTimer.PRE := 2000, [1,5].LOLOTimerSP := 2, [1,5].LOTimer.PRE := 2000, [1,5].LOTimerSP := 2, [1,5].HITimer.PRE := 2000, [1,5].HITimerSP := 2, [1,5].HIHITimer.PRE := 2000, [1,5].HIHITimerSP := 2, [1,5].EnableCfg := 1, [1,6].LOLODisable := 1, [1,6].LODisable := 1,
        [1,6].HIHIEnable := 1, [1,6].FeedPumpEnable := 1, [1,6].FeedPumpTag := 1, [1,6].HI := 6.0, [1,6].HIHI := 6.0, [1,6].PV := -0.03822385, [1,6].LOLOTimer.PRE := 2000, [1,6].LOLOTimerSP := 2, [1,6].LOTimer.PRE := 2000, [1,6].LOTimerSP := 2, [1,6].HITimer.PRE := 2000, [1,6].HITimerSP := 2, [1,6].HIHITimer.PRE := 2000, [1,6].HIHITimerSP := 2, [1,6].EnableCfg := 1, [1,7].LOLODisable := 1, [1,7].LODisable := 1, [1,7].HIHIEnable := 1, [1,7].FeedPumpEnable := 1, [1,7].FeedPumpTag := 1, [1,7].HI := 6.0, [1,7].HIHI := 6.0, [1,7].PV := -0.015335317, [1,7].LOLOTimer.PRE := 2000, [1,7].LOLOTimerSP := 2, [1,7].LOTimer.PRE := 2000, [1,7].LOTimerSP := 2, [1,7].HITimer.PRE := 2000, [1,7].HITimerSP := 2, [1,7].HIHITimer.PRE := 2000, [1,7].HIHITimerSP := 2, [1,7].EnableCfg := 1, [1,8].LOLODisable := 1, [1,8].LODisable := 1, [1,8].HIHIEnable := 1, [1,8].TransferPumpEnable := 1, [1,8].TransferPumpTag := 2, [1,8].HI := 6.0, [1,8].HIHI := 6.0, [1,8].PV := 0.014419775, [1,8].LOLOTimer.PRE := 2000, [1,8].LOLOTimerSP := 2, [1,8].LOTimer.PRE := 2000, [1,8].LOTimerSP := 2, [1,8].HITimer.PRE := 2000, [1,8].HITimerSP := 2, [1,8].HIHITimer.PRE := 2000, [1,8].HIHITimerSP := 2, [1,8].EnableCfg := 1, [1,9].Override := 1, [1,9].HI := 14.0, [1,9].HIHI := 14.0, [1,9].LOLOTimer.PRE := 2000, [1,9].LOLOTimerSP := 2, [1,9].LOTimer.PRE := 2000, [1,9].LOTimerSP := 2, [1,9].HITimer.PRE := 2000, [1,9].HITimerSP := 2, [1,9].HIHITimer.PRE := 2000, [1,9].HIHITimerSP := 2,
        [1,10].HI := 100.0, [1,10].HIHI := 100.0, [1,10].PV := 0.019073777, [1,10].LOLOTimer.PRE := 2000, [1,10].LOLOTimerSP := 2, [1,10].LOTimer.PRE := 2000, [1,10].LOTimerSP := 2, [1,10].HITimer.PRE := 2000, [1,10].HITimerSP := 2, [1,10].HIHITimer.PRE := 2000, [1,10].HIHITimerSP := 2, [1,10].EnableCfg := 1, [1,11].Override := 1, [1,11].HI := 2.0, [1,11].HIHI := 2.0, [1,11].PV := 0.0017547875, [1,11].LOLOTimer.PRE := 2000, [1,11].LOLOTimerSP := 2, [1,11].LOTimer.PRE := 2000, [1,11].LOTimerSP := 2, [1,11].HITimer.PRE := 2000, [1,11].HITimerSP := 2, [1,11].HIHITimer.PRE := 2000, [1,11].HIHITimerSP := 2, [1,11].EnableCfg := 1, [1,12].Override := 1, [1,12].HI := 2.0, [1,12].HIHI := 2.0, [1,12].PV := 0.0035858701, [1,12].LOLOTimer.PRE := 2000, [1,12].LOLOTimerSP := 2, [1,12].LOTimer.PRE := 2000, [1,12].LOTimerSP := 2, [1,12].HITimer.PRE := 2000, [1,12].HITimerSP := 2, [1,12].HIHITimer.PRE := 2000, [1,12].HIHITimerSP := 2, [1,12].EnableCfg := 1, [1,13].HI := 55.0, [1,13].HIHI := 55.0, [1,13].PV := 22.464523, [1,13].LOLOTimer.PRE := 2000, [1,13].LOLOTimerSP := 2, [1,13].LOTimer.PRE := 2000, [1,13].LOTimerSP := 2, [1,13].HITimer.PRE := 2000, [1,13].HITimerSP := 2, [1,13].HIHITimer.PRE := 2000, [1,13].HIHITimerSP := 2, [1,13].EnableCfg := 1, [1,14].Override := 1, [1,14].HI := 100.0, [1,14].HIHI := 100.0, [1,14].LOLOTimer.PRE := 1000, [1,14].LOLOTimerSP := 2, [1,14].LOTimer.PRE := 5000, [1,14].LOTimerSP := 2, [1,14].HITimer.PRE := 5000, [1,14].HITimerSP := 2, [1,14].HIHITimer.PRE := 1000,
        [1,14].HIHITimerSP := 2, [1,15].LOLODisable := 1, [1,15].LODisable := 1, [1,15].FeedPumpEnable := 1, [1,15].FeedPumpTag := 1, [1,15].HI := 60.0, [1,15].HIHI := 60.0, [1,15].PV := -0.16, [1,15].LOLOTimer.PRE := 2000, [1,15].LOLOTimerSP := 2, [1,15].LOTimer.PRE := 2000, [1,15].LOTimerSP := 2, [1,15].HITimer.PRE := 2000, [1,15].HITimerSP := 2, [1,15].HIHITimer.PRE := 2000, [1,15].HIHITimerSP := 2, [1,15].EnableCfg := 1, [1,16].Override := 1, [1,16].HI := 2.0, [1,16].HIHI := 2.0, [1,16].LOLOTimer.PRE := 2000, [1,16].LOLOTimerSP := 2, [1,16].LOTimer.PRE := 2000, [1,16].LOTimerSP := 2, [1,16].HITimer.PRE := 2000, [1,16].HITimerSP := 2, [1,16].HIHITimer.PRE := 2000, [1,16].HIHITimerSP := 2, [1,17].Override := 1, [1,17].LOLODisable := 1, [1,17].LODisable := 1, [1,17].FeedPumpEnable := 1, [1,17].TransferPumpEnable := 1, [1,17].FeedPumpTag := 1, [1,17].TransferPumpTag := 2, [1,17].HI := 15.0, [1,17].HIHI := 15.0, [1,17].LOLOTimer.PRE := 2000, [1,17].LOLOTimerSP := 2, [1,17].LOTimer.PRE := 2000, [1,17].LOTimerSP := 2, [1,17].HITimer.PRE := 2000, [1,17].HITimerSP := 2, [1,17].HIHITimer.PRE := 2000, [1,17].HIHITimerSP := 2, [1,18].Override := 1, [1,18].LOLODisable := 1, [1,18].LODisable := 1, [1,18].FeedPumpEnable := 1, [1,18].FeedPumpTag := 1, [1,18].LOLO := -1.0, [1,18].LO := -1.0, [1,18].HI := 5.0, [1,18].HIHI := 5.0, [1,18].LOLOTimer.PRE := 2000, [1,18].LOLOTimerSP := 2, [1,18].LOTimer.PRE := 2000, [1,18].LOTimerSP := 2, [1,18].HITimer.PRE := 2000, [1,18].HITimerSP := 2,
        [1,18].HIHITimer.PRE := 2000, [1,18].HIHITimerSP := 2, [1,19].Override := 1, [1,19].LOLODisable := 1, [1,19].LODisable := 1, [1,19].TransferPumpEnable := 1, [1,19].TransferPumpTag := 2, [1,19].LOLO := -1.0, [1,19].LO := -1.0, [1,19].HI := 5.0, [1,19].HIHI := 5.0, [1,19].LOLOTimer.PRE := 2000, [1,19].LOLOTimerSP := 2, [1,19].LOTimer.PRE := 2000, [1,19].LOTimerSP := 2, [1,19].HITimer.PRE := 2000, [1,19].HITimerSP := 2, [1,19].HIHITimer.PRE := 2000, [1,19].HIHITimerSP := 2, [1,20].Override := 1, [1,20].HI := 100.0, [1,20].HIHI := 100.0, [1,20].LOLOTimerSP := 2, [1,20].LOTimerSP := 2, [1,20].HITimer.EN := 1, [1,20].HITimer.DN := 1, [1,20].HITimerSP := 2, [1,20].HIHITimer.EN := 1, [1,20].HIHITimer.DN := 1, [1,20].HIHITimerSP := 2, [1,21].Override := 1, [1,21].HI := 100.0, [1,21].HIHI := 100.0, [1,21].LOLOTimerSP := 2, [1,21].LOTimerSP := 2, [1,21].HITimerSP := 2, [1,21].HIHITimerSP := 2, [1,22].Override := 1, [1,23].Override := 1, [1,24].Override := 1, [1,25].Override := 1, [1,26].Override := 1, [1,27].Override := 1, [1,28].Override := 1, [1,28].HI := 100.0, [1,28].HIHI := 100.0, [1,28].LOLOTimer.PRE := 2000, [1,28].LOLOTimerSP := 2, [1,28].LOTimer.PRE := 2000, [1,28].LOTimerSP := 2, [1,28].HITimer.PRE := 2000, [1,28].HITimerSP := 2, [1,28].HIHITimer.PRE := 2000, [1,28].HIHITimerSP := 2, [1,29].Override := 1, [1,29].HI := 100.0, [1,29].HIHI := 100.0, [1,29].LOLOTimer.PRE := 2000, [1,29].LOLOTimerSP := 2, [1,29].LOTimer.PRE := 2000,
        [1,29].LOTimerSP := 2, [1,29].HITimer.PRE := 2000, [1,29].HITimerSP := 2, [1,29].HIHITimer.PRE := 2000, [1,29].HIHITimerSP := 2, [1,30].Override := 1, [1,30].HI := 100.0, [1,30].HIHI := 100.0, [1,30].LOLOTimer.PRE := 2000, [1,30].LOLOTimerSP := 2, [1,30].LOTimer.PRE := 2000, [1,30].LOTimerSP := 2, [1,30].HITimer.PRE := 2000, [1,30].HITimerSP := 2, [1,30].HIHITimer.PRE := 2000, [1,30].HIHITimerSP := 2, [1,31].Override := 1, [1,31].HI := 100.0, [1,31].HIHI := 100.0, [1,31].LOLOTimer.PRE := 2000, [1,31].LOLOTimerSP := 2, [1,31].LOTimer.PRE := 2000, [1,31].LOTimerSP := 2, [1,31].HITimer.PRE := 2000, [1,31].HITimerSP := 2, [1,31].HIHITimer.PRE := 2000, [1,31].HIHITimerSP := 2, [1,32].Override := 1, [1,33].Override := 1, [1,34].Override := 1, [1,35].Override := 1, [1,36].Override := 1, [1,37].Override := 1, [1,38].Override := 1, [1,39].Override := 1, [1,40].LOLODisable := 1, [1,40].LODisable := 1, [1,40].FeedPumpEnable := 1, [1,40].FeedPumpTag := 1, [1,40].HI := 6.0, [1,40].HIHI := 6.0, [1,40].PV := 0.026092928, [1,40].LOLOTimer.PRE := 2000, [1,40].LOLOTimerSP := 2, [1,40].LOTimer.PRE := 2000, [1,40].LOTimerSP := 2, [1,40].HITimer.PRE := 2000, [1,40].HITimerSP := 2, [1,40].HIHITimer.PRE := 2000, [1,40].HIHITimerSP := 2, [1,40].EnableCfg := 1, [1,41].LOLODisable := 1, [1,41].LODisable := 1, [1,41].FeedPumpEnable := 1, [1,41].FeedPumpTag := 1, [1,41].HI := 6.0, [1,41].HIHI := 6.0, [1,41].PV := -0.009384299, [1,41].LOLOTimer.PRE := 2000, [1,41].LOLOTimerSP := 2,
        [1,41].LOTimer.PRE := 2000, [1,41].LOTimerSP := 2, [1,41].HITimer.PRE := 2000, [1,41].HITimerSP := 2, [1,41].HIHITimer.PRE := 2000, [1,41].HIHITimerSP := 2, [1,41].EnableCfg := 1, [1,42].LOLODisable := 1, [1,42].LODisable := 1, [1,42].FeedPumpEnable := 1, [1,42].FeedPumpTag := 1, [1,42].HI := 25.0, [1,42].HIHI := 25.0, [1,42].LOLOTimer.PRE := 2000, [1,42].LOLOTimerSP := 2, [1,42].LOTimer.PRE := 2000, [1,42].LOTimerSP := 2, [1,42].HITimer.PRE := 2000, [1,42].HITimerSP := 2, [1,42].HIHITimer.PRE := 2000, [1,42].HIHITimerSP := 2, [1,42].EnableCfg := 1, [1,43].LOLODisable := 1, [1,43].LODisable := 1, [1,43].TransferPumpEnable := 1, [1,43].TransferPumpTag := 2, [1,43].HI := 25.0, [1,43].HIHI := 25.0, [1,43].LOLOTimer.PRE := 2000, [1,43].LOLOTimerSP := 2, [1,43].LOTimer.PRE := 2000, [1,43].LOTimerSP := 2, [1,43].HITimer.PRE := 2000, [1,43].HITimerSP := 2, [1,43].HIHITimer.PRE := 2000, [1,43].HIHITimerSP := 2, [1,43].EnableCfg := 1, [1,44].LOLODisable := 1, [1,44].LODisable := 1, [1,44].FeedPumpEnable := 1, [1,44].FeedPumpTag := 1, [1,44].HI := 50.0, [1,44].HIHI := 50.0, [1,44].PV := -0.16, [1,44].LOLOTimer.PRE := 2000, [1,44].LOLOTimerSP := 2, [1,44].LOTimer.PRE := 2000, [1,44].LOTimerSP := 2, [1,44].HITimer.PRE := 2000, [1,44].HITimerSP := 2, [1,44].HIHITimer.PRE := 2000, [1,44].HIHITimerSP := 2, [1,44].EnableCfg := 1, [1,45].Override := 1, [1,45].LOLODisable := 1, [1,45].LODisable := 1, [1,45].HI := 999.0, [1,45].HIHI := 999.0, [1,45].LOLOTimer.PRE := 2000, [1,45].LOLOTimerSP := 2,
        [1,45].LOTimer.PRE := 2000, [1,45].LOTimerSP := 2, [1,45].HITimer.PRE := 2000, [1,45].HITimerSP := 2, [1,45].HIHITimer.PRE := 2000, [1,45].HIHITimerSP := 2, [1,46].Override := 1, [1,46].HI := 999.0, [1,46].HIHI := 999.0, [1,46].LOLOTimerSP := 2, [1,46].LOTimerSP := 2, [1,46].HITimerSP := 2, [1,46].HIHITimerSP := 2, [1,47].Override := 1, [1,48].Override := 1, [1,49].Override := 1, [2,0].HI := 1500.0, [2,0].HIHI := 1500.0, [2,0].LOLOTimer.PRE := 2000, [2,0].LOLOTimerSP := 2, [2,0].LOTimer.PRE := 2000, [2,0].LOTimerSP := 2, [2,0].HITimer.PRE := 2000, [2,0].HITimerSP := 2, [2,0].HIHITimer.PRE := 2000, [2,0].HIHITimerSP := 2, [2,0].EnableCfg := 1, [2,1].Override := 1, [2,1].HI := 1000.0, [2,1].HIHI := 1000.0, [2,1].PV := -12.499046, [2,1].LOLOTimer.PRE := 2000, [2,1].LOLOTimerSP := 2, [2,1].LOTimer.PRE := 2000, [2,1].LOTimerSP := 2, [2,1].HITimer.PRE := 2000, [2,1].HITimerSP := 2, [2,1].HIHITimer.PRE := 2000, [2,1].HIHITimerSP := 2, [2,2].LOLODisable := 1, [2,2].LODisable := 1, [2,2].FeedPumpEnable := 1, [2,2].FeedPumpTag := 1, [2,2].HI := 25.0, [2,2].HIHI := 25.0, [2,2].PV := -6.249523, [2,2].LOLOTimer.PRE := 2000, [2,2].LOLOTimerSP := 2, [2,2].LOTimer.PRE := 2000, [2,2].LOTimerSP := 2, [2,2].HITimer.PRE := 2000, [2,2].HITimerSP := 2, [2,2].HIHITimer.PRE := 2000, [2,2].HIHITimerSP := 2, [2,2].EnableCfg := 1, [2,3].Override := 1, [2,3].HI := 100.0, [2,3].HIHI := 100.0, [2,3].PV := -3.499525, [2,3].LOLOTimer.PRE := 1000,
        [2,3].LOLOTimerSP := 2, [2,3].LOTimer.PRE := 5000, [2,3].LOTimerSP := 2, [2,3].HITimer.PRE := 5000, [2,3].HITimerSP := 2, [2,3].HIHITimer.PRE := 1000, [2,3].HIHITimerSP := 2, [2,4].Override := 1, [2,4].HI := 100.0, [2,4].HIHI := 100.0, [2,4].PV := -24.996607, [2,4].LOLOTimer.PRE := 1000, [2,4].LOLOTimerSP := 2, [2,4].LOTimer.PRE := 5000, [2,4].LOTimerSP := 2, [2,4].HITimer.PRE := 5000, [2,4].HITimerSP := 2, [2,4].HIHITimer.PRE := 1000, [2,4].HIHITimerSP := 2, [2,5].LOLODisable := 1, [2,5].LODisable := 1, [2,5].HIHIEnable := 1, [2,5].FeedPumpEnable := 1, [2,5].FeedPumpTag := 1, [2,5].HI := 6.0, [2,5].HIHI := 6.0, [2,5].PV := -1.4998856, [2,5].LOLOTimer.PRE := 2000, [2,5].LOLOTimerSP := 2, [2,5].LOTimer.PRE := 2000, [2,5].LOTimerSP := 2, [2,5].HITimer.PRE := 2000, [2,5].HITimerSP := 2, [2,5].HIHITimer.PRE := 2000, [2,5].HIHITimerSP := 2, [2,5].EnableCfg := 1, [2,6].LOLODisable := 1, [2,6].LODisable := 1, [2,6].HIHIEnable := 1, [2,6].FeedPumpEnable := 1, [2,6].FeedPumpTag := 1, [2,6].HI := 6.0, [2,6].HIHI := 6.0, [2,6].PV := -1.4998856, [2,6].LOLOTimer.PRE := 2000, [2,6].LOLOTimerSP := 2, [2,6].LOTimer.PRE := 2000, [2,6].LOTimerSP := 2, [2,6].HITimer.PRE := 2000, [2,6].HITimerSP := 2, [2,6].HIHITimer.PRE := 2000, [2,6].HIHITimerSP := 2, [2,6].EnableCfg := 1, [2,7].LOLODisable := 1, [2,7].LODisable := 1, [2,7].HIHIEnable := 1, [2,7].FeedPumpEnable := 1, [2,7].FeedPumpTag := 1, [2,7].HI := 6.0, [2,7].HIHI := 6.0,
        [2,7].PV := -1.4998856, [2,7].LOLOTimer.PRE := 2000, [2,7].LOLOTimerSP := 2, [2,7].LOTimer.PRE := 2000, [2,7].LOTimerSP := 2, [2,7].HITimer.PRE := 2000, [2,7].HITimerSP := 2, [2,7].HIHITimer.PRE := 2000, [2,7].HIHITimerSP := 2, [2,7].EnableCfg := 1, [2,8].LOLODisable := 1, [2,8].LODisable := 1, [2,8].HIHIEnable := 1, [2,8].TransferPumpEnable := 1, [2,8].TransferPumpTag := 2, [2,8].HI := 6.0, [2,8].HIHI := 6.0, [2,8].PV := -1.4998856, [2,8].LOLOTimer.PRE := 2000, [2,8].LOLOTimerSP := 2, [2,8].LOTimer.PRE := 2000, [2,8].LOTimerSP := 2, [2,8].HITimer.PRE := 2000, [2,8].HITimerSP := 2, [2,8].HIHITimer.PRE := 2000, [2,8].HIHITimerSP := 2, [2,8].EnableCfg := 1, [2,9].Override := 1, [2,9].HI := 14.0, [2,9].HIHI := 14.0, [2,9].PV := -1.4998856, [2,9].LOLOTimer.PRE := 2000, [2,9].LOLOTimerSP := 2, [2,9].LOTimer.PRE := 2000, [2,9].LOTimerSP := 2, [2,9].HITimer.PRE := 2000, [2,9].HITimerSP := 2, [2,9].HIHITimer.PRE := 2000, [2,9].HIHITimerSP := 2, [2,10].HI := 100.0, [2,10].HIHI := 100.0, [2,10].PV := -24.998093, [2,10].LOLOTimer.PRE := 2000, [2,10].LOLOTimerSP := 2, [2,10].LOTimer.PRE := 2000, [2,10].LOTimerSP := 2, [2,10].HITimer.PRE := 2000, [2,10].HITimerSP := 2, [2,10].HIHITimer.PRE := 2000, [2,10].HIHITimerSP := 2, [2,10].EnableCfg := 1, [2,11].Override := 1, [2,11].HI := 2.0, [2,11].HIHI := 2.0, [2,11].PV := -0.49996185, [2,11].LOLOTimer.PRE := 2000, [2,11].LOLOTimerSP := 2, [2,11].LOTimer.PRE := 2000, [2,11].LOTimerSP := 2, [2,11].HITimer.PRE := 2000,
        [2,11].HITimerSP := 2, [2,11].HIHITimer.PRE := 2000, [2,11].HIHITimerSP := 2, [2,12].Override := 1, [2,12].HI := 2.0, [2,12].HIHI := 2.0, [2,12].PV := -0.49996185, [2,12].LOLOTimer.PRE := 2000, [2,12].LOLOTimerSP := 2, [2,12].LOTimer.PRE := 2000, [2,12].LOTimerSP := 2, [2,12].HITimer.PRE := 2000, [2,12].HITimerSP := 2, [2,12].HIHITimer.PRE := 2000, [2,12].HIHITimerSP := 2, [2,13].HI := 55.0, [2,13].HIHI := 55.0, [2,13].PV := -13.748952, [2,13].LOLOTimer.PRE := 2000, [2,13].LOLOTimerSP := 2, [2,13].LOTimer.PRE := 2000, [2,13].LOTimerSP := 2, [2,13].HITimer.PRE := 2000, [2,13].HITimerSP := 2, [2,13].HIHITimer.PRE := 2000, [2,13].HIHITimerSP := 2, [2,13].EnableCfg := 1, [2,14].Override := 1, [2,14].HI := 100.0, [2,14].HIHI := 100.0, [2,14].LOLOTimerSP := 2, [2,14].LOTimerSP := 2, [2,14].HITimerSP := 2, [2,14].HIHITimerSP := 2, [2,15].LOLODisable := 1, [2,15].LODisable := 1, [2,15].FeedPumpEnable := 1, [2,15].FeedPumpTag := 1, [2,15].HI := 60.0, [2,15].HIHI := 60.0, [2,15].LOLOTimer.PRE := 2000, [2,15].LOLOTimerSP := 2, [2,15].LOTimer.PRE := 2000, [2,15].LOTimerSP := 2, [2,15].HITimer.PRE := 2000, [2,15].HITimerSP := 2, [2,15].HIHITimer.PRE := 2000, [2,15].HIHITimerSP := 2, [2,15].EnableCfg := 1, [2,16].Override := 1, [2,16].PV := -0.4999322, [2,16].LOLOTimerSP := 2, [2,16].LOTimerSP := 2, [2,16].HITimerSP := 2, [2,16].HIHITimerSP := 2, [2,17].Override := 1, [2,17].PV := -2.499796, [2,17].LOLOTimerSP := 2, [2,17].LOTimerSP := 2, [2,17].HITimerSP := 2,
        [2,17].HIHITimerSP := 2, [2,18].Override := 1, [2,18].PV := -2.499796, [2,18].LOLOTimerSP := 2, [2,18].LOTimerSP := 2, [2,18].HITimerSP := 2, [2,18].HIHITimerSP := 2, [2,19].Override := 1, [2,19].PV := -2.499796, [2,19].LOLOTimerSP := 2, [2,19].LOTimerSP := 2, [2,19].HITimerSP := 2, [2,19].HIHITimerSP := 2, [2,20].Override := 1, [2,20].PV := 100.0, [2,20].LOLOTimerSP := 2, [2,20].LOTimerSP := 2, [2,20].HITimer.EN := 1, [2,20].HITimer.DN := 1, [2,20].HITimerSP := 2, [2,20].HIHITimer.EN := 1, [2,20].HIHITimer.DN := 1, [2,20].HIHITimerSP := 2, [2,21].Override := 1, [2,21].LOLOTimerSP := 2, [2,21].LOTimerSP := 2, [2,21].HITimerSP := 2, [2,21].HIHITimerSP := 2, [2,22].Override := 1, [2,22].PV := 0.5047684, [2,23].Override := 1, [2,23].PV := 0.1161975, [2,24].Override := 1, [2,24].PV := 0.16, [2,25].Override := 1, [2,25].PV := -0.3333333, [2,26].Override := 1, [2,26].PV := 63.88032, [2,27].Override := 1, [2,27].PV := -37.40687, [2,28].Override := 1, [2,28].HI := 100.0, [2,28].HIHI := 100.0, [2,28].PV := 22.8542, [2,28].LOLOTimer.PRE := 2000, [2,28].LOLOTimerSP := 2, [2,28].LOTimer.PRE := 2000, [2,28].LOTimerSP := 2, [2,28].HITimer.PRE := 2000, [2,28].HITimerSP := 2, [2,28].HIHITimer.PRE := 2000, [2,28].HIHITimerSP := 2, [2,29].Override := 1, [2,29].HI := 100.0, [2,29].HIHI := 100.0, [2,29].PV := 21.877623, [2,29].LOLOTimer.PRE := 2000, [2,29].LOLOTimerSP := 2, [2,29].LOTimer.PRE := 2000, [2,29].LOTimerSP := 2,
        [2,29].HITimer.PRE := 2000, [2,29].HITimerSP := 2, [2,29].HIHITimer.PRE := 2000, [2,29].HIHITimerSP := 2, [2,30].Override := 1, [2,30].HI := 100.0, [2,30].HIHI := 100.0, [2,30].PV := 21.877623, [2,30].LOLOTimer.PRE := 2000, [2,30].LOLOTimerSP := 2, [2,30].LOTimer.PRE := 2000, [2,30].LOTimerSP := 2, [2,30].HITimer.PRE := 2000, [2,30].HITimerSP := 2, [2,30].HIHITimer.PRE := 2000, [2,30].HIHITimerSP := 2, [2,31].Override := 1, [2,31].HI := 100.0, [2,31].HIHI := 100.0, [2,31].PV := 21.877623, [2,31].LOLOTimer.PRE := 2000, [2,31].LOLOTimerSP := 2, [2,31].LOTimer.PRE := 2000, [2,31].LOTimerSP := 2, [2,31].HITimer.PRE := 2000, [2,31].HITimerSP := 2, [2,31].HIHITimer.PRE := 2000, [2,31].HIHITimerSP := 2, [2,32].Override := 1, [2,32].PV := 0.1837702, [2,33].Override := 1, [2,33].PV := -0.6615715, [2,34].Override := 1, [2,34].PV := 0.6615715, [2,35].Override := 1, [2,35].PV := 222.0, [2,36].Override := 1, [2,37].Override := 1, [2,37].PV := -0.03181506, [2,38].Override := 1, [2,39].Override := 1, [2,40].LOLODisable := 1, [2,40].LODisable := 1, [2,40].FeedPumpEnable := 1, [2,40].FeedPumpTag := 1, [2,40].HI := 6.0, [2,40].HIHI := 6.0, [2,40].LOLOTimer.PRE := 2000, [2,40].LOLOTimerSP := 2, [2,40].LOTimer.PRE := 2000, [2,40].LOTimerSP := 2, [2,40].HITimer.PRE := 2000, [2,40].HITimerSP := 2, [2,40].HIHITimer.PRE := 2000, [2,40].HIHITimerSP := 2, [2,40].EnableCfg := 1, [2,41].LOLODisable := 1, [2,41].LODisable := 1, [2,41].FeedPumpEnable := 1, [2,41].FeedPumpTag := 1,
        [2,41].HI := 6.0, [2,41].HIHI := 6.0, [2,41].LOLOTimer.PRE := 2000, [2,41].LOLOTimerSP := 2, [2,41].LOTimer.PRE := 2000, [2,41].LOTimerSP := 2, [2,41].HITimer.PRE := 2000, [2,41].HITimerSP := 2, [2,41].HIHITimer.PRE := 2000, [2,41].HIHITimerSP := 2, [2,41].EnableCfg := 1, [2,42].LOLODisable := 1, [2,42].LODisable := 1, [2,42].FeedPumpEnable := 1, [2,42].FeedPumpTag := 1, [2,42].HI := 45.0, [2,42].HIHI := 45.0, [2,42].LOLOTimer.PRE := 2000, [2,42].LOLOTimerSP := 2, [2,42].LOTimer.PRE := 2000, [2,42].LOTimerSP := 2, [2,42].HITimer.PRE := 2000, [2,42].HITimerSP := 2, [2,42].HIHITimer.PRE := 2000, [2,42].HIHITimerSP := 2, [2,42].EnableCfg := 1, [2,43].LOLODisable := 1, [2,43].LODisable := 1, [2,43].TransferPumpEnable := 1, [2,43].TransferPumpTag := 2, [2,43].HI := 25.0, [2,43].HIHI := 25.0, [2,43].LOLOTimer.PRE := 2000, [2,43].LOLOTimerSP := 2, [2,43].LOTimer.PRE := 2000, [2,43].LOTimerSP := 2, [2,43].HITimer.PRE := 2000, [2,43].HITimerSP := 2, [2,43].HIHITimer.PRE := 2000, [2,43].HIHITimerSP := 2, [2,43].EnableCfg := 1, [2,44].LOLODisable := 1, [2,44].LODisable := 1, [2,44].FeedPumpEnable := 1, [2,44].FeedPumpTag := 1, [2,44].HI := 50.0, [2,44].HIHI := 50.0, [2,44].LOLOTimer.PRE := 2000, [2,44].LOLOTimerSP := 2, [2,44].LOTimer.PRE := 2000, [2,44].LOTimerSP := 2, [2,44].HITimer.PRE := 2000, [2,44].HITimerSP := 2, [2,44].HIHITimer.PRE := 2000, [2,44].HIHITimerSP := 2, [2,44].EnableCfg := 1, [2,45].Override := 1, [2,45].HI := 999.0, [2,45].HIHI := 999.0, [2,45].LOLOTimerSP := 2,
        [2,45].LOTimerSP := 2, [2,45].HITimerSP := 2, [2,45].HIHITimerSP := 2, [2,46].Override := 1, [2,46].HI := 999.0, [2,46].HIHI := 999.0, [2,46].LOLOTimerSP := 2, [2,46].LOTimerSP := 2, [2,46].HITimerSP := 2, [2,46].HIHITimerSP := 2, [2,47].Override := 1, [2,48].Override := 1, [2,49].Override := 1, [3,1].PV := -0.06111238, [3,1].EnableCfg := 1, [3,2].PV := -0.03822385, [3,2].EnableCfg := 1, [3,3].HIAlarm := 1, [3,3].HIHIAlarm := 1, [3,3].HIAlarmONS := 1, [3,3].HIHIAlarmONS := 1, [3,3].Value := 4, [3,3].ValueHMI := 4, [3,3].PV := 0.2228261, [3,3].HITimer.EN := 1, [3,3].HITimer.DN := 1, [3,3].HIHITimer.EN := 1, [3,3].HIHITimer.DN := 1, [3,3].EnableCfg := 1, [3,4].PV := -0.03387503, [3,4].EnableCfg := 1, [3,5].HIAlarm := 1, [3,5].HIHIAlarm := 1, [3,5].HIAlarmONS := 1, [3,5].HIHIAlarmONS := 1, [3,5].Value := 4, [3,5].ValueHMI := 4, [3,5].PV := 1.033333, [3,5].HITimer.EN := 1, [3,5].HITimer.DN := 1, [3,5].HIHITimer.EN := 1, [3,5].HIHITimer.DN := 1, [3,5].EnableCfg := 1, [3,6].EnableCfg := 1, [3,7].EnableCfg := 1, [3,8].PV := -25.10109, [3,8].EnableCfg := 1, [3,9].LOLODisable := 1, [3,9].LODisable := 1, [3,9].FeedPumpEnable := 1, [3,9].TransferPumpEnable := 1, [3,9].FeedPumpTag := 1, [3,9].TransferPumpTag := 2, [3,9].EnableCfg := 1, [3,10].HIAlarm := 1, [3,10].HIHIAlarm := 1, [3,10].LOLODisable := 1, [3,10].LODisable := 1, [3,10].FeedPumpEnable := 1, [3,10].HIAlarmONS := 1,
